(* IEC 61131-3 sources: SortJet_MasterSPS_Aufbau.fbsproj/07_Auftragsverwaltung/BasisSchrittketten, 22 files *)

(* ---- Shuttle_Austransport.fb.st ---- *)
(* METADATA
{
	"v3Meta": {
		"objectGuid": "ac2be6b1-afec-449b-a8c9-7faca61891b0"
	}
}
*)
FUNCTION_BLOCK Shuttle_Austransport
VAR_INPUT

  // BOOLEAN
  bpReset                : BOOL;

  // WORD
  wStation               : WORD;
  wWand                  : WORD;

  // STRUKTUR
  Auftragsdaten          : Auftragsdaten_ST;

END_VAR
VAR_OUTPUT

  // BOOLEAN
  bpDone                 : BOOL;
  bpFehler               : BOOL;

END_VAR
VAR

  // BOOLEAN
  blStationQuittiertScheiben : BOOL;

  // WORD
  wlAustransportstation  : WORD;

  // INT
  ilScheibenZuQuittieren : INT;

  // STEPS
  steplSchritt           : STEPS_TE;

END_VAR
//-------------------------------------------------------------------------------------------------
// STEUERUNG AUSTRANSPORT
//-------------------------------------------------------------------------------------------------
IF ( Auftragsdaten.wAuftrag = eStation_Austransport) THEN

  CASE steplSchritt OF

    // AUSTRANSPORT ===============================================
    STEP_0_E:
      (* Hinweis:
         - Ueberpruefung des Sicherheitskreises
      *)
      IF checkSafetyCircuitsNotBlocked(starrShuttleBasisParameter[wStation]) AND NOT bgShuttleAustransportSperren[wStation]  THEN
        steplSchritt := STEP_10_E;
      END_IF

    // AUSTRANSPORT ===============================================
    STEP_10_E:
      // Auftragsdaten pruefen:
      //  - Sollte es fehler in der Auftragsdatenstruktur geben wird in den Fehlerschritt 900
      //    gesprungen. Die Fehlerauswertung findet in der Funktion Shuttledaten_Pruefen statt.
      steplSchritt := STEP_20_E;

      IF NOT AuftragsdatenPruefen( wStation, wWand, Auftragsdaten) THEN
        steplSchritt := STEP_900_E;
      END_IF

    // AUSTRANSPORT ===============================================
    STEP_20_E:
      // ---------------------------------------------------------------------------------------
      //  AUSTRANSPORT BEDINGUNGEN PRUEFEN
      //
      //  Hinweis:
      // - n/c
      // ---------------------------------------------------------------------------------------

      (* Hinweis:
         - Uebergabe der Quellstation [Sender] fuer den Austransport [Zum ueberpruefen des Zustandes der Station]
      *)
      wlAustransportstation := Auftragsdaten.wTransferstationsNr1;

      starrShuttleBasisParameter[wStation].bRueckwaertsTransportieren[wWand] := FALSE;
      starrShuttleBasisParameter[wStation].bTransferstationTransfershuttle[wWand] := FALSE;

      (* Hinweis:
         - Auftragsdaten ans Shuttle übergeben
      *)
      ilScheibenZuQuittieren :=WORD_TO_INT( Auftragsdaten.wAnzahlScheiben);

      (* Hinweis:
         - Auftragsdaten uebergeben
      *)
      starrShuttleBasisParameter[wStation].pAuftrag[wWand] := Auftragsdaten;

      (* Hinweis:
         - Scheibenführung / Wandverstellung anstellen
         - Aus dem Speicher: Speicherslot dicke nehmen ; von einer Station die Scheibendicke nehmen
      *)
      IF ( starrShuttleBasisParameter[wStation].pAuftrag[wWand].rAuftragsDicke <= wgMKScheibenDicke13mm ) THEN
        starrShuttleBasisParameter[wStation].pAuftrag[wWand].stAuftragsOptionen.eDickenverstellung    := eZylinderStellung16mm;
      ELSIF ( starrShuttleBasisParameter[wStation].pAuftrag[wWand].rAuftragsDicke <= wgMKScheibenDicke19mm ) THEN
        starrShuttleBasisParameter[wStation].pAuftrag[wWand].stAuftragsOptionen.eDickenverstellung    := eZylinderStellung23mm;
      ELSIF ( starrShuttleBasisParameter[wStation].pAuftrag[wWand].rAuftragsDicke <= wgMKScheibenDicke24mm ) THEN
        starrShuttleBasisParameter[wStation].pAuftrag[wWand].stAuftragsOptionen.eDickenverstellung    := eZylinderStellung29mm;
      END_IF

      // Kippen
      starrShuttleBasisParameter[wStation].pAuftrag[wWand].stAuftragsOptionen.eKippen_SollPosition                  := starrShuttleBasisParameter[wStation].stMKs.stSchnittstellendaten.aAustransporte.Kippen[wlAustransportstation];
      starrShuttleBasisParameter[wStation].pAuftrag[wWand].stAuftragsOptionen.eKippen_SollPosition_NachEintransport := 0;
      starrShuttleBasisParameter[wStation].pAuftrag[wWand].stAuftragsOptionen.eKippen_SollPosition_NachAustransport := starrShuttleBasisParameter[wStation].stMKs.stSchnittstellendaten.aAustransporte.KippenNachAustransport[wlAustransportstation];

      // Hub
      starrShuttleBasisParameter[wStation].pAuftrag[wWand].stAuftragsOptionen.eHub                  := starrShuttleBasisParameter[wStation].stMKs.stSchnittstellendaten.aAustransporte.Hub[wlAustransportstation];
      starrShuttleBasisParameter[wStation].pAuftrag[wWand].stAuftragsOptionen.eHub_NachEintransport := 0;
      starrShuttleBasisParameter[wStation].pAuftrag[wWand].stAuftragsOptionen.eHub_NachAustransport := starrShuttleBasisParameter[wStation].stMKs.stSchnittstellendaten.aAustransporte.HubNachAustransport[wlAustransportstation];

      // Greifer [Ausbaustufe stStationsAufbau.bGreifer]: Greiferseite je Partnerstation, Zangenoeffnung wie die Scheibenfuehrung
      starrShuttleBasisParameter[wStation].pAuftrag[wWand].stAuftragsOptionen.eGreiferTyp   := eGreiferDefault;
      IF ( starrShuttleBasisParameter[wStation].stMKs.stStationsAufbau.bGreifer[wWand] ) THEN
        starrShuttleBasisParameter[wStation].pAuftrag[wWand].stAuftragsOptionen.eGreiferTyp := starrShuttleBasisParameter[wStation].stMKs.stSchnittstellendaten.aAustransporte.Greifer[wlAustransportstation];
      END_IF
      starrShuttleBasisParameter[wStation].pAuftrag[wWand].stAuftragsOptionen.eGreiferZangeStellung := starrShuttleBasisParameter[wStation].pAuftrag[wWand].stAuftragsOptionen.eDickenverstellung;

      // Scheibentyp prüfen
      starrShuttleBasisParameter[wStation].wGlasTyp[wWand] := eScheibe_Default;
      IF ( Auftragsdaten.rAuftragsLaenge >= starrShuttleBasisParameter[wStation].stMKs.stStationsParameter.rLaengeUebergroesseScheibe ) THEN
        starrShuttleBasisParameter[wStation].wGlasTyp[wWand] := eScheibe_Maximal;
      END_IF

      (* Hinweis:
         - Stations-Zustand pruefen
      *)
      CASE wlAustransportstation OF

        // Transfershuttles
        cERSTES_TRANSFERSHUTTLE..cLETZTES_TRANSFERSHUTTLE:
          steplSchritt := STEP_200_E;

        // Stationen
        cERSTE_STATION..cLETZTE_STATION:
          IF ( ( Job_Stationen.AuftragsdatenWand[wlAustransportstation, Auftragsdaten.wTransferwand].wAuftrag = eStation_Kein_Auftrag )
               OR ( Job_Stationen.AuftragsdatenWand[wlAustransportstation, Auftragsdaten.wTransferwand].wAuftrag = eStation_Belegt )
               OR ( Job_Stationen.AuftragsdatenWand[wlAustransportstation, Auftragsdaten.wTransferwand].wAuftrag = eStation_Durchtransport ) )
          THEN
            steplSchritt := STEP_100_E;
          END_IF

        cERSTE_FREMDANLAGE_AUSLAUF..cLETZTE_FREMDANLAGE_AUSLAUF:
          IF ( Auftragsdaten.wTransferstationsNr2 <> 0 ) THEN
            IF   ( Job_Fremdanlage.AuftragsdatenFremdanlage[wlAustransportstation].wAuftrag = eStation_Kein_Auftrag )
                 AND ( Job_Stationen.AuftragsdatenWand[Auftragsdaten.wTransferstationsNr2, Auftragsdaten.wTransferwand].wAuftrag = eStation_Kein_Auftrag )
            THEN
              steplSchritt := STEP_100_E;
            END_IF
          ELSE
            IF ( Job_Fremdanlage.AuftragsdatenFremdanlage[wlAustransportstation].wAuftrag = eStation_Kein_Auftrag )
            THEN
              steplSchritt := STEP_100_E;
            END_IF
          END_IF

        // Fremdanlage
        cERSTE_FREMDANLAGE_EINLAUF..cLETZTE_FREMDANLAGE_EINLAUF:
          ;

        // Faecherwagen direkt (Transferstation 1): nur mit dem Greifer. Ohne Greifer geht es in den Faecherwagen ueber ein
        // Transfershuttle mit bTransferShuttleFuerFaecherwagen (Transferstation 1 = Transfershuttle, Transferstation 2 = Faecherwagen)
        cERSTE_FAECHERWAGENSTATIONS_NR..cLETZTE_FAECHERWAGENSTATIONS_NR:
          IF ( starrShuttleBasisParameter[wStation].pAuftrag[wWand].stAuftragsOptionen.eGreiferTyp <> eGreiferDefault ) THEN
            IF ( starrFaecherwagenBasisParameter[wlAustransportstation].OutGlasTransport[cWAND_1].bBereitZumEintransport ) THEN
              steplSchritt := STEP_100_E;
            END_IF
          ELSE
            wpgFehlerdaten[0] := starrShuttleBasisParameter[wStation].stMKs.stStationsNummern.NummerExtern;
            wpgFehlerdaten[1] := wWand;
            SpsError( eFehler_Station,
                      cMELDUNG_AUFTRAGSDATEN_FALSCHE_AUSLAUFSTATION,
                      starrShuttleBasisParameter[wStation].stMKs.stStationsNummern.NummerIntern,
                      AutomatikkreisBestimmen(starrShuttleBasisParameter[wStation].stMKs.stStationsNummern.NummerSPS),
                      wpgFehlerdaten );

            steplSchritt := STEP_900_E;
          END_IF

        ELSE
          wpgFehlerdaten[0] := starrShuttleBasisParameter[wStation].stMKs.stStationsNummern.NummerExtern;
          wpgFehlerdaten[1] := wWand;
          SpsError( eFehler_Station,
                    cMELDUNG_AUFTRAGSDATEN_FALSCHE_AUSLAUFSTATION,
                    starrShuttleBasisParameter[wStation].stMKs.stStationsNummern.NummerIntern,
                    AutomatikkreisBestimmen(starrShuttleBasisParameter[wStation].stMKs.stStationsNummern.NummerSPS),
                    wpgFehlerdaten );

          steplSchritt := STEP_900_E;

      END_CASE

    // AUSTRANSPORT ==============================================
    STEP_100_E:
      (* Hinweis:
         - Auftrag ab Station übergeben und Shuttle Informationen zuweisen
      *)
      CASE wlAustransportstation OF

        // Stationen
        cERSTE_STATION..cLETZTE_STATION:

          IF AutomatikAktiv(wlAustransportstation) THEN

            (* Hinweis:
               - Auftragsdaten in Transferstation kopieren
            *)
            IF NOT ( Job_Stationen.AuftragsdatenWand[wlAustransportstation, Auftragsdaten.wTransferwand].wAuftrag = eStation_Durchtransport ) THEN
              Job_Stationen.AuftragsdatenWand[wlAustransportstation, Auftragsdaten.wTransferwand]           := AuftragsdatenUmkopieren(FALSE, FALSE, Auftragsdaten);
              Job_Stationen.AuftragsdatenWand[wlAustransportstation, Auftragsdaten.wTransferwand].wAuftrag  := eStation_Eintransport;
            END_IF

            (* Hinweis:
               - Kopplung zur Transferstation herstellen
            *)
            starrShuttleBasisParameter[wStation].InGlasTransportNachfolger[wWand] := starrStationBasisParameter[wlAustransportstation].OutGlasTransport[Auftragsdaten.wTransferwand];
            starrShuttleBasisParameter[wStation].InGlasTransportVorgaenger[wWand] := starrStationBasisParameter[wlAustransportstation].OutGlasTransport[Auftragsdaten.wTransferwand];

            (* Hinweis:
               - Daten an das Shuttle uebergeben
            *)
            starrShuttleBasisParameter[wStation].bAustransport[wWand]                  := TRUE;
            starrShuttleBasisParameter[wStation].bRueckwaertsTransportieren[wWand]     := ( starrShuttleBasisParameter[wStation].stMKs.stSchnittstellendaten.aAustransporte.Station[wlAustransportstation] = Rueckwaertig );

            steplSchritt := STEP_400_E;

          END_IF

        cERSTE_FREMDANLAGE_AUSLAUF..cLETZTE_FREMDANLAGE_AUSLAUF:

          IF ( Auftragsdaten.wTransferstationsNr2 <> 0 ) THEN

            IF AutomatikAktiv(Auftragsdaten.wTransferstationsNr2) THEN

              (* Hinweis:
                 - Kopplung zur Transferstation herstellen
              *)
              starrShuttleBasisParameter[wStation].InGlasTransportNachfolger[wWand] := starrStationBasisParameter[Auftragsdaten.wTransferstationsNr2].OutGlasTransport[Auftragsdaten.wTransferwand];
              starrShuttleBasisParameter[wStation].InGlasTransportVorgaenger[wWand] := starrStationBasisParameter[Auftragsdaten.wTransferstationsNr2].OutGlasTransport[Auftragsdaten.wTransferwand];

              (* Hinweis:
                 - Auftragsdaten in Transferstation kopieren
              *)
              Job_Fremdanlage.AuftragsdatenFremdanlage[wlAustransportstation]          := AuftragsdatenUmkopieren(FALSE, FALSE, Auftragsdaten);
              Job_Fremdanlage.AuftragsdatenFremdanlage[wlAustransportstation].wAuftrag := eStation_Eintransport;

              (* Hinweis:
                 - Daten an das Shuttle uebergeben
              *)
              starrShuttleBasisParameter[wStation].bAustransport[wWand]                  := TRUE;
              starrShuttleBasisParameter[wStation].bRueckwaertsTransportieren[wWand]     := ( starrShuttleBasisParameter[wStation].stMKs.stSchnittstellendaten.aAustransporte.Station[wlAustransportstation] = Rueckwaertig );

              steplSchritt := STEP_400_E;

            END_IF

          ELSE

            (* Hinweis:
               - Kopplung zur Transferstation herstellen
            *)
            starrShuttleBasisParameter[wStation].InGlasTransportNachfolger[wWand] := starrFremdanlageAuslaufStationBasisParameter[wlAustransportstation].OutGlasTransport[cWAND_1];
            starrShuttleBasisParameter[wStation].InGlasTransportVorgaenger[wWand] := starrFremdanlageAuslaufStationBasisParameter[wlAustransportstation].OutGlasTransport[cWAND_1];
            starrFremdanlageAuslaufStationBasisParameter[wlAustransportstation].InGlasTransportVorgaenger[cWAND_1] :=  starrShuttleBasisParameter[wStation].OutGlasTransport[wWand];

            (* Hinweis:
               - Auftragsdaten in Transferstation kopieren
            *)
            Job_Fremdanlage.AuftragsdatenFremdanlage[wlAustransportstation]          := AuftragsdatenUmkopieren(FALSE, FALSE, Auftragsdaten);
            Job_Fremdanlage.AuftragsdatenFremdanlage[wlAustransportstation].wAuftrag := eStation_Eintransport;

            (* Hinweis:
               - Daten an das Shuttle uebergeben
            *)
            starrShuttleBasisParameter[wStation].bAustransport[wWand]              := TRUE;
            starrShuttleBasisParameter[wStation].bRueckwaertsTransportieren[wWand] := ( starrShuttleBasisParameter[wStation].stMKs.stSchnittstellendaten.aAustransporte.Station[wlAustransportstation] = Rueckwaertig );

            steplSchritt := STEP_400_E;

          END_IF

        cERSTE_FAECHERWAGENSTATIONS_NR..cLETZTE_FAECHERWAGENSTATIONS_NR:
          (* Hinweis:
             - Austransport in den Faecherwagen mit dem Greifer (Greiferseite im Auftrag)
          *)
          starrShuttleBasisParameter[wStation].bRueckwaertsTransportieren[wWand] := FALSE;
          starrShuttleBasisParameter[wStation].bAustransport[wWand]              := TRUE;

          steplSchritt := STEP_400_E;

      END_CASE

    // AUSTRANSPORT ===============================================
    STEP_200_E:
      // ---------------------------------------------------------------------------------------
      //  EINTRANSPORT MITTELS TRANSFERSHUTTLE
      //
      //  Hinweis:
      //  - Transferstation2 = 0   => Eintransport mit nur einem Transfershuttle
      //  - Transferstation2 <> 0  => Eintransport im Transfershuttle-Verbund
      // ---------------------------------------------------------------------------------------

      IF ( Auftragsdaten.wTransferstationsNr2 = 0 OR starrTransfershuttleBasisParameter[wlAustransportstation].stMKs.stStationsOptionen.stTransfershuttle.bTransferShuttleFuerFaecherwagen ) THEN

        IF (  ( Job_Shuttle.AuftragsdatenTransfershuttle[wlAustransportstation].wAuftrag = eStation_Kein_Auftrag ) ) THEN
          steplSchritt := STEP_210_E;
        END_IF

      ELSE
        VailiderenTransfershuttleVerbund ( wTransferstation1 := wlAustransportstation,
                                           wTransferstation2 := Auftragsdaten.wTransferstationsNr2 );

        IF (  ( Job_Shuttle.AuftragsdatenTransfershuttle[wlAustransportstation].wAuftrag = eStation_Kein_Auftrag )
             AND ( Job_Shuttle.AuftragsdatenTransfershuttle[Auftragsdaten.wTransferstationsNr2].wAuftrag  = eStation_Kein_Auftrag ) )
        THEN
          steplSchritt := STEP_220_E;
        END_IF

      END_IF

    // AUSTRANSPORT ===============================================
    STEP_210_E:
      // ---------------------------------------------------------------------------------------
      //  EINTRANSPORT TRANSFERSHUTTLE [DEFAULT]
      //
      //  Hinweis:
      // - n/c
      // ---------------------------------------------------------------------------------------

      (* Hinweis:
         - Kopplung
      *)
      IF ( starrShuttleBasisParameter[wStation].stMKs.stSchnittstellendaten.aAustransporte.Station[wlAustransportstation] = Rueckwaertig ) THEN
        starrTransfershuttleBasisParameter[wlAustransportstation].InGlasTransportNachfolger[wWand] := starrShuttleBasisParameter[wStation].OutGlasTransport[wWand];
        starrShuttleBasisParameter[wStation].InGlasTransportVorgaenger[wWand] := starrTransfershuttleBasisParameter[wlAustransportstation].OutGlasTransport[wWand];

      ELSE
        starrTransfershuttleBasisParameter[wlAustransportstation].InGlasTransportVorgaenger[wWand] := starrShuttleBasisParameter[wStation].OutGlasTransport[wWand];
        starrShuttleBasisParameter[wStation].InGlasTransportNachfolger[wWand] := starrTransfershuttleBasisParameter[wlAustransportstation].OutGlasTransport[wWand];

      END_IF

      (* Hinweis:
         - TS auf FW koppeln
      *)
      IF   starrTransfershuttleBasisParameter[wlAustransportstation].stMKs.stStationsOptionen.stTransfershuttle.bTransferShuttleFuerFaecherwagen
           AND IsBetweenWORD(Auftragsdaten.wTransferstationsNr2, cERSTE_FAECHERWAGENSTATIONS_NR, cLETZTE_FAECHERWAGENSTATIONS_NR)
      THEN
        IF ( starrShuttleBasisParameter[wStation].stMKs.stSchnittstellendaten.aAustransporte.Station[wlAustransportstation] = Rueckwaertig ) THEN
          starrTransfershuttleBasisParameter[wlAustransportstation].InGlasTransportVorgaenger[wWand] := starrFaecherwagenBasisParameter[Auftragsdaten.wTransferstationsNr2].OutGlasTransport[cWAND_1];
        ELSE
          starrTransfershuttleBasisParameter[wlAustransportstation].InGlasTransportNachfolger[wWand] := starrFaecherwagenBasisParameter[Auftragsdaten.wTransferstationsNr2].OutGlasTransport[cWAND_1];
        END_IF
      END_IF

      (* Hinweis:
         - Neuen Auftag in den FIFO [Warteschlange] eintragen
      *)
      Job_Shuttle.AuftragsdatenTransfershuttle[wlAustransportstation]          := AuftragsdatenUmkopieren(FALSE, FALSE, Auftragsdaten);
      Job_Shuttle.AuftragsdatenTransfershuttle[wlAustransportstation].wAuftrag := eStation_Eintransport;

      starrShuttleBasisParameter[wStation].bScheibentrennen[wWand]                := FALSE;
      starrShuttleBasisParameter[wStation].bRueckwaertsTransportieren[wWand]      := ( starrShuttleBasisParameter[wStation].stMKs.stSchnittstellendaten.aAustransporte.Station[wlAustransportstation] = Rueckwaertig );
      starrShuttleBasisParameter[wStation].bAustransport[wWand]                   := TRUE;
      starrShuttleBasisParameter[wStation].bTransferstationTransfershuttle[wWand] := TRUE;

      steplSchritt := STEP_400_E;

    // AUSTRANSPORT ===============================================
    STEP_220_E:
      // ---------------------------------------------------------------------------------------
      //  EINTRANSPORT TRANSFERSHUTTLE [VERBUND]
      //
      //  Hinweis:
      //  - n/c
      // ---------------------------------------------------------------------------------------

      (* Hinweis:
         - Kopplung
      *)
      IF ( starrShuttleBasisParameter[wStation].stMKs.eStationsTyp = eInputshuttle ) THEN
        starrTransfershuttleBasisParameter[wlAustransportstation].InGlasTransportVorgaenger[wWand] := starrShuttleBasisParameter[wStation].OutGlasTransport[wWand];
        starrShuttleBasisParameter[wStation].InGlasTransportNachfolger[wWand] := starrTransfershuttleBasisParameter[wlAustransportstation].OutGlasTransport[wWand];

      ELSE
        starrTransfershuttleBasisParameter[wlAustransportstation].InGlasTransportNachfolger[wWand] := starrShuttleBasisParameter[wStation].OutGlasTransport[wWand];
        starrShuttleBasisParameter[wStation].InGlasTransportVorgaenger[wWand] := starrTransfershuttleBasisParameter[wlAustransportstation].OutGlasTransport[wWand];

      END_IF

      (* Hinweis:
         - Transfershuttle koppeln
      *)
      aTransfershuttles[wlAustransportstation].stpInTransportVerbund  := aTransfershuttles[Auftragsdaten.wTransferstationsNr2].stpOutTransportVerbund;
      aTransfershuttles[Auftragsdaten.wTransferstationsNr2].stpInTransportVerbund   := aTransfershuttles[wlAustransportstation].stpOutTransportVerbund;

      (* Hinweis:
         - Auftragsdaten an die Transfershuttle uebergeben
      *)
      Job_Shuttle.AuftragsdatenTransfershuttle[wlAustransportstation]          := AuftragsdatenUmkopieren(FALSE, FALSE, Auftragsdaten);
      Job_Shuttle.AuftragsdatenTransfershuttle[wlAustransportstation].wAuftrag := eStation_Eintransport;

      Job_Shuttle.AuftragsdatenTransfershuttle[Auftragsdaten.wTransferstationsNr2]           := AuftragsdatenUmkopieren(TRUE, FALSE, Auftragsdaten);
      Job_Shuttle.AuftragsdatenTransfershuttle[Auftragsdaten.wTransferstationsNr2].wAuftrag  := eStation_Transportkopplung;

      starrShuttleBasisParameter[wStation].bScheibentrennen[wWand]                := FALSE;
      starrShuttleBasisParameter[wStation].bRueckwaertsTransportieren[wWand]      := ( starrShuttleBasisParameter[wStation].stMKs.stSchnittstellendaten.aAustransporte.Station[wlAustransportstation] = Rueckwaertig );
      starrShuttleBasisParameter[wStation].bAustransport[wWand]                   := TRUE;
      starrShuttleBasisParameter[wStation].bTransferstationTransfershuttle[wWand] := TRUE;

      steplSchritt := STEP_400_E;

    // AUSTRANSPORT ===============================================
    STEP_400_E:
      // ---------------------------------------------------------------------------------------
      //  QUITTIERUNGEN UND EINTRANSPORT- ABSCHLUSS
      //
      //  Hinweis:
      //  - Scheibenquittieren: Message zur MMI
      // ---------------------------------------------------------------------------------------
      blStationQuittiertScheiben := starrShuttleBasisParameter[wStation].stMKs.stSchnittstellendaten.aAustransporte.bStationQuittiertScheibe[wlAustransportstation];

      IF ( starrShuttleBasisParameter[wStation].OutGlasTransport[wWand].bQuittScheibe ) THEN

        IF ( ilScheibenZuQuittieren > 0 ) THEN

          wSps2MmiZielStation  := Auftragsdaten.wTransferstationsNr1;
          wSps2MmiQuellStation := starrShuttleBasisParameter[wStation].stMKs.stStationsNummern.NummerIntern;
          wSps2MmiZielWand     := Auftragsdaten.wTransferwand;
          wSps2MmiQuellWand    := wWand;
          dwSps2MmiWartezeit   := starrShuttleBasisParameter[wStation].dwWartezeit[wWand];
          wSPS2MMIAuftragstyp  := 1;

          MsgToMmi(auftragsnr_w := SB0_SPS_QUIT_SHEET_ORDER );
        END_IF

        ilScheibenZuQuittieren := ilScheibenZuQuittieren - 1;

      END_IF

      (* Hinweis:
         - Abschliessen des Austransports
      *)
      IF ( starrShuttleBasisParameter[wStation].bAustransportAbgeschlossen[wWand] ) THEN

        starrShuttleBasisParameter[wStation].bAustransport[wWand]                 := FALSE;
        starrShuttleBasisParameter[wStation].bRueckwaertsTransportieren[wWand]    := FALSE;

        steplSchritt := STEP_410_E;
      END_IF

      (* Fehlerbehandlung:
         - Inputshuttle
      *)
      IF ( starrShuttleBasisParameter[wStation].bFehler ) THEN
        SpsError( eFehler_Station,
                  starrShuttleBasisParameter[wStation].wFehlerNummer,
                  starrShuttleBasisParameter[wStation].stMKs.stStationsNummern.NummerIntern,
                  AutomatikkreisBestimmen(starrShuttleBasisParameter[wStation].stMKs.stStationsNummern.NummerSPS),
                  starrShuttleBasisParameter[wStation].awFehlerInformationen );

        steplSchritt := STEP_900_E;
      END_IF

    // AUSTRANSPORT ==============================================
    STEP_410_E:
      (* Anmerkung:
         - Gueltige Anzahl von Scheiben wurden quittiert
      *)
      IF ( ilScheibenZuQuittieren = 0 ) THEN
        steplSchritt := STEP_1000_E;

      (* Anmerkung:
         - Zu wenig Scheiben quittiert
      *)
      ELSIF ( ilScheibenZuQuittieren > 0 ) THEN
        wpgFehlerdaten[0] := starrShuttleBasisParameter[wStation].stMKs.stStationsNummern.NummerExtern;
        wpgFehlerdaten[1] := wWand;

        SpsError( eFehler_Station,
                  cMELDUNG_STATION_ZUWENIG_SCHEIBEN_QUITTIERT_WAND_AUSTRANSPORT,
                  starrShuttleBasisParameter[wStation].stMKs.stStationsNummern.NummerIntern,
                  AutomatikkreisBestimmen(starrShuttleBasisParameter[wStation].stMKs.stStationsNummern.NummerSPS),
                  wpgFehlerdaten );

        steplSchritt := STEP_900_E;

      (* Anmerkung:
         - Zu viele Scheiben quittiert
      *)
      ELSIF ( ilScheibenZuQuittieren < 0 ) THEN
        wpgFehlerdaten[0] := starrShuttleBasisParameter[wStation].stMKs.stStationsNummern.NummerExtern;
        wpgFehlerdaten[1] := wWand;

        SpsError( eFehler_Station,
                  cMELDUNG_STATION_ZUVIELE_SCHEIBEN_QUITTIERT_WAND_AUSTRANSPORT,
                  starrShuttleBasisParameter[wStation].stMKs.stStationsNummern.NummerIntern,
                  AutomatikkreisBestimmen(starrShuttleBasisParameter[wStation].stMKs.stStationsNummern.NummerSPS),
                  wpgFehlerdaten );

        steplSchritt := STEP_900_E;
      END_IF

    // AUSTRANSPORT ===============================================
    STEP_900_E:
      bpFehler := TRUE;

    // AUSTRANSPORT ===============================================
    STEP_1000_E:
      bpDone := TRUE;
      Auftragsdaten.wAuftrag := eStation_Kein_Auftrag;

  // AUSTRANSPORT ===============================================
  END_CASE

END_IF

IF bpReset THEN
  bpFehler := FALSE;
  bpDone := FALSE;
  bpReset := FALSE;
  starrShuttleBasisParameter[wStation].bAustransport[wWand] := FALSE;
  starrShuttleBasisParameter[wStation].bTransferstationTransfershuttle[wWand] := FALSE;
  steplSchritt := STEP_0_E;
END_IF
END_FUNCTION_BLOCK

(* ---- Shuttle_Durchtransport.fb.st ---- *)
(* METADATA
{
	"v3Meta": {
		"objectGuid": "d20ae107-ce5b-4166-b2bd-9e4de3a442ef"
	}
}
*)
FUNCTION_BLOCK Shuttle_Durchtransport
VAR_INPUT

  // BOOLEAN
  bpReset                : BOOL;

  // WORD
  wStation               : WORD;
  wWand                  : WORD;

  // STRUKTUR
  Auftragsdaten          : Auftragsdaten_ST;

END_VAR
VAR_OUTPUT

  // BOOLEAN
  bpDone                 : BOOL;
  bpFehler               : BOOL;

END_VAR
VAR

  // BOOLEAN
  blStationQuittiertScheiben             : BOOL;
  blKopplungGefundenEintransport         : BOOL;
  blKopplungGefundenAustransport         : BOOL;

  // WORD
  wlEintransportstation : WORD;
  wlAustransportstation : WORD;

  // INT
  ilScheibenZuQuittieren : INT;

  // STEPS
  steplSchritt           : STEPS_TE;

END_VAR

//-------------------------------------------------------------------------------------------------
// STEUERUNG DURCHTRANSPORT
//-------------------------------------------------------------------------------------------------
IF Auftragsdaten.wAuftrag = eStation_Durchtransport THEN
  CASE steplSchritt OF
    // DURCHTRANSPORT =================================
    STEP_0_E:
      (* Hinweis:
         - Ueberpruefung des Sicherheitskreises
      *)
      IF checkSafetyCircuitsNotBlocked(starrShuttleBasisParameter[wStation]) AND NOT bgShuttleEintransportSperren[wStation] AND NOT bgShuttleAustransportSperren[wStation]  THEN
        steplSchritt := STEP_10_E;
      END_IF

    // DURCHTRANSPORT ==================================================
    STEP_10_E:
      // Auftragsdaten pruefen:
      //  - Sollte es fehler in der Auftragsdatenstruktur geben wird in den Fehlerschritt 900
      //    gesprungen. Die Fehlerauswertung findet in der Funktion Shuttledaten_Pruefen statt.
      steplSchritt := STEP_20_E;

      IF NOT AuftragsdatenPruefen( wStation, wWand, Auftragsdaten) THEN
        steplSchritt := STEP_900_E;
      END_IF

    // DURCHTRANSPORT =================================
    STEP_20_E:
      (* Hinweis:
         - Kopplung fuer diesen Auftrag neu bestimmen. Sonst ueberschreibt ein Merker aus dem letzten Auftrag den Fehlerschritt.
      *)
      blKopplungGefundenEintransport := FALSE;
      blKopplungGefundenAustransport := FALSE;

      (* Hinweis:
         - Uebergabe der Quellstation [Sender] fuer den Austransport [Zum ueberpruefen des Zustandes der Station]
      *)
      wlEintransportstation := Auftragsdaten.wTransferstationsNr1;
      wlAustransportstation := Auftragsdaten.wTransferstationsNr2;

      (* Hinweis:
         - Zuweisung Transportkopplung
      *)
      CASE wlEintransportstation OF

        // Stationen
        cERSTE_STATION..cLETZTE_STATION:
          (* Hinweis:
             - Transportkopplung
          *)
          IF ( starrShuttleBasisParameter[wStation].stMKs.stSchnittstellendaten.aEintransporte.Station[wlEintransportstation] = Vorwaertig ) THEN
            starrShuttleBasisParameter[wStation].InGlasTransportVorgaenger[wWand] := starrStationBasisParameter[wlEintransportstation].OutGlasTransport[Auftragsdaten.wTransferwand];
          ELSE
            starrShuttleBasisParameter[wStation].InGlasTransportNachfolger[wWand] := starrStationBasisParameter[wlEintransportstation].OutGlasTransport[Auftragsdaten.wTransferwand];
          END_IF
          blKopplungGefundenEintransport := TRUE;

        ELSE
          wpgFehlerdaten[0] := starrShuttleBasisParameter[wStation].stMKs.stStationsNummern.NummerExtern;
          wpgFehlerdaten[1] := wlEintransportstation;
          SpsError( eFehler_Station,
                    cMELDUNG_AUFTRAGSDATEN_FALSCHE_EINLAUFSTATION,
                    starrShuttleBasisParameter[wStation].stMKs.stStationsNummern.NummerIntern,
                    AutomatikkreisBestimmen(starrShuttleBasisParameter[wStation].stMKs.stStationsNummern.NummerSPS),
                    wpgFehlerdaten );

          steplSchritt := STEP_900_E;

      END_CASE

      (* Hinweis:
         - Zuweisung Transportkopplung
      *)
      CASE wlAustransportstation OF

        // Stationen
        cERSTE_STATION..cLETZTE_STATION:
          (* Hinweis:
             - Transportkopplung
          *)
          IF ( starrShuttleBasisParameter[wStation].stMKs.stSchnittstellendaten.aAustransporte.Station[wlAustransportstation] = Vorwaertig ) THEN
            starrShuttleBasisParameter[wStation].InGlasTransportNachfolger[wWand] := starrStationBasisParameter[wlAustransportstation].OutGlasTransport[Auftragsdaten.wTransferwand];
          ELSE
            starrShuttleBasisParameter[wStation].InGlasTransportVorgaenger[wWand] := starrStationBasisParameter[wlAustransportstation].OutGlasTransport[Auftragsdaten.wTransferwand];
          END_IF
          blKopplungGefundenAustransport := TRUE;

        cERSTE_FREMDANLAGE_AUSLAUF..cLETZTE_FREMDANLAGE_AUSLAUF:
          (* Hinweis:
             - Transportkopplung
          *)
          IF ( starrShuttleBasisParameter[wStation].stMKs.stSchnittstellendaten.aAustransporte.Station[wlAustransportstation] = Vorwaertig ) THEN
            starrShuttleBasisParameter[wStation].InGlasTransportNachfolger[wWand] := starrFremdanlageAuslaufStationBasisParameter[wlAustransportstation].OutGlasTransport[cWAND_1];
          ELSE
            starrShuttleBasisParameter[wStation].InGlasTransportVorgaenger[wWand] := starrFremdanlageAuslaufStationBasisParameter[wlAustransportstation].OutGlasTransport[cWAND_1];
          END_IF
          blKopplungGefundenAustransport := TRUE;

        ELSE
          wpgFehlerdaten[0] := starrShuttleBasisParameter[wStation].stMKs.stStationsNummern.NummerExtern;
          wpgFehlerdaten[1] := wlAustransportstation;
          SpsError( eFehler_Station,
                    cMELDUNG_AUFTRAGSDATEN_FALSCHE_AUSLAUFSTATION,
                    starrShuttleBasisParameter[wStation].stMKs.stStationsNummern.NummerIntern,
                    AutomatikkreisBestimmen(starrShuttleBasisParameter[wStation].stMKs.stStationsNummern.NummerSPS),
                    wpgFehlerdaten );

          steplSchritt := STEP_900_E;

      END_CASE

      IF blKopplungGefundenEintransport AND blKopplungGefundenAustransport THEN
        steplSchritt := STEP_30_E;
      END_IF

    // DURCHTRANSPORT =================================
    STEP_30_E:

      (* Hinweis:
         - Scheibenquittierung
      *)
      ilScheibenZuQuittieren := WORD_TO_INT(Auftragsdaten.wAnzahlScheiben);

      (* Hinweis:
         - Auftrags- Optionen bestimmen und zuweisen
      *)
      Auftragsdaten.stAuftragsOptionen.eKippen_SollPosition := starrShuttleBasisParameter[wStation].stMKs.stSchnittstellendaten.aEintransporte.Kippen[wlEintransportstation];

      IF ( Auftragsdaten.rAuftragsDicke < wgUnterteilerMinMaxGlasdicke ) THEN
        Auftragsdaten.stAuftragsOptionen.eDickenverstellung := eZylinderStellung16mm;
      ELSE
        Auftragsdaten.stAuftragsOptionen.eDickenverstellung := eZylinderStellung23mm;
      END_IF
      Auftragsdaten.stAuftragsOptionen.eDrehen_Sollposition := 0;
      Auftragsdaten.stAuftragsOptionen.eDrehen_Sollposition_NachAustransport := 0;
      Auftragsdaten.stAuftragsOptionen.eKippen_SollPosition_NachAustransport := 0;
      Auftragsdaten.stAuftragsOptionen.eGlastransport := 0;
      Auftragsdaten.stAuftragsOptionen.eHub                  := starrShuttleBasisParameter[wStation].stMKs.stSchnittstellendaten.aEintransporte.Hub[wlEintransportstation];
      Auftragsdaten.stAuftragsOptionen.eHub_NachEintransport := 0;
      Auftragsdaten.stAuftragsOptionen.eHub_NachAustransport := 0;
      Auftragsdaten.stAuftragsOptionen.eQuerachse := 0;
      Auftragsdaten.stAuftragsOptionen.eAchsrichtung := 0;
      Auftragsdaten.stAuftragsOptionen.wMaxTransportGeschwindigkeit:= 0;
      Auftragsdaten.stAuftragsOptionen.eDrehen_Sollposition_NachEintransport := 0;
      Auftragsdaten.stAuftragsOptionen.eKippen_SollPosition_NachEintransport := 0;

      (* Hinweis:
         - Auftragsdaten zuweisen und Eintransport der Station starten
      *)
      starrShuttleBasisParameter[wStation].pAuftrag[wWand] := Auftragsdaten;

      starrShuttleBasisParameter[wStation].bScheibentrennen[wWand]           := FALSE;
      starrShuttleBasisParameter[wStation].bRueckwaertsTransportieren[wWand] := ( starrShuttleBasisParameter[wStation].stMKs.stSchnittstellendaten.aEintransporte.Station[wlEintransportstation] = Rueckwaertig )
                                                                                AND ( starrShuttleBasisParameter[wStation].stMKs.stSchnittstellendaten.aAustransporte.Station[wlAustransportstation] = Rueckwaertig );
      starrShuttleBasisParameter[wStation].bDurchtransport[wWand]            := TRUE;

      steplSchritt := STEP_40_E;

    // AUSTRANSPORT =================================
    STEP_40_E:

      (* Hinweis:
         - Scheibenzaehler dekrementieren
         - Scheibe quittieren, sofern dies nötig ist
      *)
      blStationQuittiertScheiben := starrShuttleBasisParameter[wStation].stMKs.stSchnittstellendaten.aEintransporte.bStationQuittiertScheibe[wlEintransportstation];

      IF ( starrShuttleBasisParameter[wStation].OutGlasTransport[wWand].bQuittScheibe ) THEN

        IF ( ilScheibenZuQuittieren > 0 ) AND blStationQuittiertScheiben THEN

          wSps2MmiZielStation  := starrShuttleBasisParameter[wStation].stMKs.stStationsNummern.NummerIntern;
          wSps2MmiQuellStation := wlEintransportstation;
          wSps2MmiZielWand     := Auftragsdaten.wStationsWand;
          wSps2MmiQuellWand    := Auftragsdaten.wTransferwand;
          dwSps2MmiWartezeit   := starrShuttleBasisParameter[wStation].dwWartezeit[wWand];
          wSPS2MMIAuftragstyp  := 0;

          MsgToMmi(auftragsnr_w := SB0_SPS_QUIT_SHEET_ORDER );

        END_IF

        ilScheibenZuQuittieren := ilScheibenZuQuittieren - 1;

      END_IF

      (* Hinweis:
         - Abschliessen des Austransport
      *)
      IF ( starrShuttleBasisParameter[wStation].bDurchtransportAbgeschlossen[wWand] ) THEN
        starrShuttleBasisParameter[wStation].bRueckwaertsTransportieren[wWand] := FALSE;
        starrShuttleBasisParameter[wStation].bDurchtransport[wWand] := FALSE;
        steplSchritt := STEP_1000_E;
      END_IF

      (* Fehlerbehandlung:
         - Station
      *)
      IF ( starrShuttleBasisParameter[wStation].bFehler ) THEN
        SpsError( eFehler_Station,
                  starrShuttleBasisParameter[wStation].wFehlerNummer,
                  starrShuttleBasisParameter[wStation].stMKs.stStationsNummern.NummerIntern,
                  AutomatikkreisBestimmen(starrShuttleBasisParameter[wStation].stMKs.stStationsNummern.NummerSPS),
                  starrShuttleBasisParameter[wStation].awFehlerInformationen );

        starrShuttleBasisParameter[wStation].bDurchtransport[wWand] := FALSE;
        starrShuttleBasisParameter[wStation].bRueckwaertsTransportieren[wWand] := FALSE;
        steplSchritt := STEP_900_E;
      END_IF

    // DURCHTRANSPORT =================================
    STEP_900_E:
      bpFehler := TRUE;

    // DURCHTRANSPORT =================================
    STEP_1000_E:
      bpDone := TRUE;
      Auftragsdaten.wAuftrag := eStation_Kein_Auftrag;

  END_CASE

END_IF

IF bpReset THEN
  bpFehler := FALSE;
  bpReset := FALSE;
  bpDone := FALSE;
  blKopplungGefundenEintransport := FALSE;
  blKopplungGefundenAustransport := FALSE;
  steplSchritt := STEP_0_E;
  starrShuttleBasisParameter[wStation].bRueckwaertsTransportieren[wWand] := FALSE;
  starrShuttleBasisParameter[wStation].bDurchtransport[wWand] := FALSE;
END_IF
END_FUNCTION_BLOCK

(* ---- Shuttle_Eintransport.fb.st ---- *)
(* METADATA
{
	"v3Meta": {
		"objectGuid": "07a4896b-4b10-421b-8c15-d73c62ab9e42"
	}
}
*)
FUNCTION_BLOCK Shuttle_Eintransport
VAR_INPUT

  // BOOLEAN
  bpReset                : BOOL;

  // WORD
  wStation               : WORD;
  wWand                  : WORD;

  // STRUKTUR
  Auftragsdaten          : Auftragsdaten_ST;

END_VAR
VAR_OUTPUT

  // BOOLEAN
  bpDone                 : BOOL;
  bpFehler               : BOOL;

END_VAR
VAR

  // BOOLEAN
  blStationQuittiertScheiben : BOOL;

  // WORD
  wlEintransportstation  : WORD;

  // INT
  ilScheibenZuQuittieren : INT;

  // STEPS
  steplSchritt           : STEPS_TE;

END_VAR

//-------------------------------------------------------------------------------------------------
// STEUERUNG EINTRANSPORT
//-------------------------------------------------------------------------------------------------
IF ( Auftragsdaten.wAuftrag = eStation_Eintransport ) THEN

  CASE steplSchritt OF

    // EINTRANSPORT ==============================================
    STEP_0_E:
      (* Hinweis:
         - Ueberpruefung des Sicherheitskreises
      *)
      IF checkSafetyCircuitsNotBlocked(starrShuttleBasisParameter[wStation]) AND NOT bgShuttleEintransportSperren[wStation] THEN
        steplSchritt := STEP_10_E;
      END_IF

    // EINTRANSPORT ==============================================
    STEP_10_E:
      // Auftragsdaten pruefen:
      //   - Sollte es fehler in der Auftragsdatenstruktur geben wird in den Fehlerschritt 900
      //   - gesprungen. Die Fehlerauswertung findet in der Funktion Shuttledaten_Pruefen statt.
      steplSchritt := STEP_20_E;

      IF NOT AuftragsdatenPruefen( wStation, wWand, Auftragsdaten) THEN
        steplSchritt := STEP_900_E;
      END_IF

    // EINTRANSPORT ==============================================
    STEP_20_E:
      (* Hinweis:
         - Uebergabe der Quellstation [Sender] fuer den Austransport [Zum ueberpruefen des Zustandes der Station]
      *)
      wlEintransportstation := Auftragsdaten.wTransferstationsNr1;

      starrShuttleBasisParameter[wStation].bRueckwaertsTransportieren[wWand] := FALSE;
      starrShuttleBasisParameter[wStation].bTransferstationTransfershuttle[wWand] := FALSE;

      (* Hinweis:
         - Auftragsdaten ans Shuttle übergeben
      *)
      ilScheibenZuQuittieren := WORD_TO_INT( Auftragsdaten.wAnzahlScheiben );

      (* Hinweis:
         - Auftragsdaten uebergeben
      *)
      starrShuttleBasisParameter[wStation].pAuftrag[wWand] := Auftragsdaten;

      (* Hinweis:
         - Scheibenführung / Wandverstellung anstellen
         - Aus dem Speicher: Speicherslot dicke nehmen ; von einer Station die Scheibendicke nehmen
      *)
      IF ( starrShuttleBasisParameter[wStation].pAuftrag[wWand].rAuftragsDicke <= wgMKScheibenDicke13mm ) THEN
        starrShuttleBasisParameter[wStation].pAuftrag[wWand].stAuftragsOptionen.eDickenverstellung    := eZylinderStellung16mm;
      ELSIF ( starrShuttleBasisParameter[wStation].pAuftrag[wWand].rAuftragsDicke <= wgMKScheibenDicke19mm ) THEN
        starrShuttleBasisParameter[wStation].pAuftrag[wWand].stAuftragsOptionen.eDickenverstellung    := eZylinderStellung23mm;
      ELSIF ( starrShuttleBasisParameter[wStation].pAuftrag[wWand].rAuftragsDicke <= wgMKScheibenDicke24mm ) THEN
        starrShuttleBasisParameter[wStation].pAuftrag[wWand].stAuftragsOptionen.eDickenverstellung    := eZylinderStellung29mm;
      END_IF

      // Kippen
      starrShuttleBasisParameter[wStation].pAuftrag[wWand].stAuftragsOptionen.eKippen_SollPosition                  := starrShuttleBasisParameter[wStation].stMKs.stSchnittstellendaten.aEintransporte.Kippen[Auftragsdaten.wTransferstationsNr1];
      starrShuttleBasisParameter[wStation].pAuftrag[wWand].stAuftragsOptionen.eKippen_SollPosition_NachEintransport := starrShuttleBasisParameter[wStation].stMKs.stSchnittstellendaten.aEintransporte.KippenNachEintransport[Auftragsdaten.wTransferstationsNr1];
      starrShuttleBasisParameter[wStation].pAuftrag[wWand].stAuftragsOptionen.eKippen_SollPosition_NachAustransport := 0;

      // Hub
      starrShuttleBasisParameter[wStation].pAuftrag[wWand].stAuftragsOptionen.eHub                  := starrShuttleBasisParameter[wStation].stMKs.stSchnittstellendaten.aEintransporte.Hub[Auftragsdaten.wTransferstationsNr1];
      starrShuttleBasisParameter[wStation].pAuftrag[wWand].stAuftragsOptionen.eHub_NachEintransport := starrShuttleBasisParameter[wStation].stMKs.stSchnittstellendaten.aEintransporte.HubNachEintransport[Auftragsdaten.wTransferstationsNr1];
      starrShuttleBasisParameter[wStation].pAuftrag[wWand].stAuftragsOptionen.eHub_NachAustransport := 0;

      // Glastransport
      starrShuttleBasisParameter[wStation].pAuftrag[wWand].stAuftragsOptionen.eGlastransport := starrShuttleBasisParameter[wStation].stMKs.stSchnittstellendaten.aEintransporte.Glastransport[Auftragsdaten.wTransferstationsNr1];

      // Greifer [Ausbaustufe stStationsAufbau.bGreifer]: Greiferseite je Partnerstation, Zangenoeffnung wie die Scheibenfuehrung
      starrShuttleBasisParameter[wStation].pAuftrag[wWand].stAuftragsOptionen.eGreiferTyp := eGreiferDefault;
      IF ( starrShuttleBasisParameter[wStation].stMKs.stStationsAufbau.bGreifer[wWand] ) THEN
        starrShuttleBasisParameter[wStation].pAuftrag[wWand].stAuftragsOptionen.eGreiferTyp := starrShuttleBasisParameter[wStation].stMKs.stSchnittstellendaten.aEintransporte.Greifer[Auftragsdaten.wTransferstationsNr1];
      END_IF
      starrShuttleBasisParameter[wStation].pAuftrag[wWand].stAuftragsOptionen.eGreiferZangeStellung := starrShuttleBasisParameter[wStation].pAuftrag[wWand].stAuftragsOptionen.eDickenverstellung;

      // Scheibentyp prüfen
      starrShuttleBasisParameter[wStation].wGlasTyp[wWand] := eScheibe_Default;
      IF ( Auftragsdaten.rAuftragsLaenge >= starrShuttleBasisParameter[wStation].stMKs.stStationsParameter.rLaengeUebergroesseScheibe ) THEN
        starrShuttleBasisParameter[wStation].wGlasTyp[wWand] := eScheibe_Maximal;
      END_IF

      (* Anmerkung:
         - Zielstation abfragen ob diese bereit sind zum Austransport
           => Status der Glas-Sender Station pruefen
      *)
      CASE wlEintransportstation OF

        // Shuttles
        cERSTES_SHUTTLE..cLETZTES_SHUTTLE: // ... macht wenig Sinn
          ;

        // Transfershuttles
        cERSTES_TRANSFERSHUTTLE..cLETZTES_TRANSFERSHUTTLE:
          steplSchritt := STEP_200_E;

        // Stationen
        cERSTE_STATION..cLETZTE_STATION:
          IF ( ( Job_Stationen.AuftragsdatenWand[wlEintransportstation, Auftragsdaten.wTransferwand].wAuftrag = eStation_Warte_Auf_Austransport )
               OR ( Job_Stationen.AuftragsdatenWand[wlEintransportstation, Auftragsdaten.wTransferwand].wAuftrag = eStation_Belegt ) )
          THEN
            steplSchritt := STEP_100_E;
          END_IF

        cERSTE_FREMDANLAGE_AUSLAUF..cLETZTE_FREMDANLAGE_AUSLAUF:
          ;

        cERSTE_FREMDANLAGE_EINLAUF..cLETZTE_FREMDANLAGE_EINLAUF:
          ;

        // Faecherwagen direkt (Transferstation 1): nur mit dem Greifer. Ohne Greifer geht es aus dem Faecherwagen ueber ein
        // Transfershuttle mit bTransferShuttleFuerFaecherwagen (Transferstation 1 = Transfershuttle, Transferstation 2 = Faecherwagen)
        cERSTE_FAECHERWAGENSTATIONS_NR..cLETZTE_FAECHERWAGENSTATIONS_NR:
          IF ( starrShuttleBasisParameter[wStation].pAuftrag[wWand].stAuftragsOptionen.eGreiferTyp <> eGreiferDefault ) THEN
            IF ( starrFaecherwagenBasisParameter[wlEintransportstation].OutGlasTransport[cWAND_1].bBereitZumAustransport ) THEN
              steplSchritt := STEP_100_E;
            END_IF
          ELSE
            wpgFehlerdaten[0] := starrShuttleBasisParameter[wStation].stMKs.stStationsNummern.NummerExtern;
            wpgFehlerdaten[1] := wlEintransportstation;
            SpsError( eFehler_Station,
                      cMELDUNG_AUFTRAGSDATEN_FALSCHE_EINLAUFSTATION,
                      starrShuttleBasisParameter[wStation].stMKs.stStationsNummern.NummerIntern,
                      AutomatikkreisBestimmen(wStation),
                      wpgFehlerdaten );

            steplSchritt := STEP_900_E;
          END_IF

        ELSE
          wpgFehlerdaten[0] := starrShuttleBasisParameter[wStation].stMKs.stStationsNummern.NummerExtern;
          wpgFehlerdaten[1] := wlEintransportstation;
          SpsError( eFehler_Station,
                    cMELDUNG_AUFTRAGSDATEN_FALSCHE_EINLAUFSTATION,
                    starrShuttleBasisParameter[wStation].stMKs.stStationsNummern.NummerIntern,
                    AutomatikkreisBestimmen(wStation),
                    wpgFehlerdaten );

          steplSchritt := STEP_900_E;

      END_CASE

    // EINTRANSPORT ==============================================
    STEP_100_E:
      // ---------------------------------------------------------------------------------------
      //  EINTRANSPORT MITTELS STATIONEN [RKT, SF, ETC.]
      //
      //  Hinweis:
      // - n/c
      // ---------------------------------------------------------------------------------------

      (* Anmerkung:
         - Starten des Eintransports [Glas-Empfaenger]
         - Initiieren des  des Austransports [Glas-Empfaenger]
      *)
      CASE wlEintransportstation OF

        cERSTE_STATION..cLETZTE_STATION:

          IF AutomatikAktiv(wlEintransportstation) THEN

            (* Hinweis:
               - Auftragsdaten in Transferstation kopieren
            *)
            Job_Stationen.AuftragsdatenWand[wlEintransportstation, Auftragsdaten.wTransferwand]           := AuftragsdatenUmkopieren(FALSE, FALSE, Auftragsdaten);
            Job_Stationen.AuftragsdatenWand[wlEintransportstation, Auftragsdaten.wTransferwand].wAuftrag  := eStation_Austransport;

            (* Hinweis:
               - Kopplung zur Transferstation herstellen
            *)
            starrShuttleBasisParameter[wStation].InGlasTransportVorgaenger[wWand] := starrStationBasisParameter[wlEintransportstation].OutGlasTransport[Auftragsdaten.wTransferwand];
            starrShuttleBasisParameter[wStation].InGlasTransportNachfolger[wWand] := starrStationBasisParameter[wlEintransportstation].OutGlasTransport[Auftragsdaten.wTransferwand];

            (* Hinweis:
               - Starten des Eintransports
            *)
            starrShuttleBasisParameter[wStation].bScheibentrennen[wWand] := NOT Auftragsdaten.stAuftragsInformationen.cBIT_SRC_WALL_1_EMPTY;
            starrShuttleBasisParameter[wStation].bRueckwaertsTransportieren[wWand] := ( starrShuttleBasisParameter[wStation].stMKs.stSchnittstellendaten.aEintransporte.Station[wlEintransportstation] = Rueckwaertig );
            starrShuttleBasisParameter[wStation].bEintransport[wWand] := TRUE;

            steplSchritt := STEP_400_E;

          END_IF

        cERSTE_FREMDANLAGE_AUSLAUF..cLETZTE_FREMDANLAGE_AUSLAUF:
          ;

        cERSTE_FREMDANLAGE_EINLAUF..cLETZTE_FREMDANLAGE_EINLAUF:
          ;

        cERSTE_FAECHERWAGENSTATIONS_NR..cLETZTE_FAECHERWAGENSTATIONS_NR:
          (* Hinweis:
             - Eintransport aus dem Faecherwagen mit dem Greifer (Greiferseite im Auftrag)
          *)
          starrShuttleBasisParameter[wStation].bScheibentrennen[wWand]           := FALSE;
          starrShuttleBasisParameter[wStation].bRueckwaertsTransportieren[wWand] := FALSE;
          starrShuttleBasisParameter[wStation].bEintransport[wWand]              := TRUE;

          steplSchritt := STEP_400_E;

      END_CASE

    // EINTRANSPORT ==============================================
    STEP_200_E:
      // ---------------------------------------------------------------------------------------
      //  EINTRANSPORT MITTELS TRANSFERSHUTTLE
      //
      //  Hinweis:
      //  - Transferstation2 = 0   => Eintransport mit nur einem Transfershuttle
      //  - Transferstation2 <> 0  => Eintransport im Transfershuttle-Verbund
      // ---------------------------------------------------------------------------------------

      IF ( Auftragsdaten.wTransferstationsNr2 = 0 OR starrTransfershuttleBasisParameter[wlEintransportstation].stMKs.stStationsOptionen.stTransfershuttle.bTransferShuttleFuerFaecherwagen ) THEN

        IF (  ( Job_Shuttle.AuftragsdatenTransfershuttle[wlEintransportstation].wAuftrag = eStation_Kein_Auftrag ) ) THEN
          steplSchritt := STEP_210_E;
        END_IF

      ELSE
        VailiderenTransfershuttleVerbund ( wTransferstation1 := wlEintransportstation,
                                           wTransferstation2 := Auftragsdaten.wTransferstationsNr2 );

        IF (  ( Job_Shuttle.AuftragsdatenTransfershuttle[wlEintransportstation].wAuftrag = eStation_Kein_Auftrag )
             AND ( Job_Shuttle.AuftragsdatenTransfershuttle[Auftragsdaten.wTransferstationsNr2].wAuftrag  = eStation_Kein_Auftrag ) )
        THEN
          steplSchritt := STEP_220_E;
        END_IF

      END_IF

    // EINTRANSPORT ==============================================
    STEP_210_E:
      // ---------------------------------------------------------------------------------------
      //  EINTRANSPORT TRANSFERSHUTTLE [DEFAULT]
      //
      //  Hinweis:
      // - n/c
      // ---------------------------------------------------------------------------------------

      (* Hinweis:
         - Kopplung
      *)
      IF ( starrShuttleBasisParameter[wStation].stMKs.stSchnittstellendaten.aEintransporte.Station[wlEintransportstation] = Rueckwaertig ) THEN
        starrTransfershuttleBasisParameter[wlEintransportstation].InGlasTransportVorgaenger[wWand] := starrShuttleBasisParameter[wStation].OutGlasTransport[wWand];
        starrShuttleBasisParameter[wStation].InGlasTransportNachfolger[wWand] := starrTransfershuttleBasisParameter[wlEintransportstation].OutGlasTransport[wWand];

      ELSE
        starrTransfershuttleBasisParameter[wlEintransportstation].InGlasTransportNachfolger[wWand] := starrShuttleBasisParameter[wStation].OutGlasTransport[wWand];
        starrShuttleBasisParameter[wStation].InGlasTransportVorgaenger[wWand] := starrTransfershuttleBasisParameter[wlEintransportstation].OutGlasTransport[wWand];

      END_IF

      (* Hinweis:
         - TS auf FW koppeln
      *)
      IF   starrTransfershuttleBasisParameter[wlEintransportstation].stMKs.stStationsOptionen.stTransfershuttle.bTransferShuttleFuerFaecherwagen
           AND IsBetweenWORD(Auftragsdaten.wTransferstationsNr2, cERSTE_FAECHERWAGENSTATIONS_NR, cLETZTE_FAECHERWAGENSTATIONS_NR)
      THEN
        IF ( starrShuttleBasisParameter[wStation].stMKs.stSchnittstellendaten.aEintransporte.Station[wlEintransportstation] = Rueckwaertig ) THEN
          starrTransfershuttleBasisParameter[wlEintransportstation].InGlasTransportNachfolger[wWand] := starrFaecherwagenBasisParameter[Auftragsdaten.wTransferstationsNr2].OutGlasTransport[cWAND_1];
        ELSE
          starrTransfershuttleBasisParameter[wlEintransportstation].InGlasTransportVorgaenger[wWand] := starrFaecherwagenBasisParameter[Auftragsdaten.wTransferstationsNr2].OutGlasTransport[cWAND_1];
        END_IF
      END_IF

      (* Hinweis:
         - Neuen Auftag in den FIFO [Warteschlange] eintragen
      *)
      Job_Shuttle.AuftragsdatenTransfershuttle[wlEintransportstation]          := AuftragsdatenUmkopieren(FALSE, FALSE, Auftragsdaten);
      Job_Shuttle.AuftragsdatenTransfershuttle[wlEintransportstation].wAuftrag := eStation_Austransport;

      starrShuttleBasisParameter[wStation].bScheibentrennen[wWand]                := FALSE;
      starrShuttleBasisParameter[wStation].bRueckwaertsTransportieren[wWand]      := ( starrShuttleBasisParameter[wStation].stMKs.stSchnittstellendaten.aEintransporte.Station[wlEintransportstation] = Rueckwaertig );
      starrShuttleBasisParameter[wStation].bEintransport[wWand]                   := TRUE;
      starrShuttleBasisParameter[wStation].bTransferstationTransfershuttle[wWand] := TRUE;

      steplSchritt := STEP_400_E;

    // EINTRANSPORT ==============================================
    STEP_220_E:
      // ---------------------------------------------------------------------------------------
      //  EINTRANSPORT TRANSFERSHUTTLE [VERBUND]
      //
      //  Hinweis:
      //  - n/c
      // ---------------------------------------------------------------------------------------

      (* Hinweis:
         - Kopplung
      *)
      IF ( starrShuttleBasisParameter[wStation].stMKs.eStationsTyp = eInputshuttle ) THEN
        starrTransfershuttleBasisParameter[wlEintransportstation].InGlasTransportVorgaenger[cWAND_1] := starrShuttleBasisParameter[wStation].OutGlasTransport[wWand];
        starrShuttleBasisParameter[wStation].InGlasTransportNachfolger[wWand] := starrTransfershuttleBasisParameter[wlEintransportstation].OutGlasTransport[cWAND_1];

      ELSE
        starrTransfershuttleBasisParameter[wlEintransportstation].InGlasTransportNachfolger[cWAND_1] := starrShuttleBasisParameter[wStation].OutGlasTransport[wWand];
        starrShuttleBasisParameter[wStation].InGlasTransportVorgaenger[wWand] := starrTransfershuttleBasisParameter[wlEintransportstation].OutGlasTransport[cWAND_1];

      END_IF

      (* Hinweis:
         - Transfershuttle koppeln
      *)
      aTransfershuttles[wlEintransportstation].stpInTransportVerbund := aTransfershuttles[Auftragsdaten.wTransferstationsNr2].stpOutTransportVerbund;
      aTransfershuttles[Auftragsdaten.wTransferstationsNr2].stpInTransportVerbund  := aTransfershuttles[wlEintransportstation].stpOutTransportVerbund;

      (* Hinweis:
         - Auftragsdaten an die Transfershuttle uebergeben
      *)
      Job_Shuttle.AuftragsdatenTransfershuttle[wlEintransportstation]            := AuftragsdatenUmkopieren(FALSE, FALSE, Auftragsdaten);
      Job_Shuttle.AuftragsdatenTransfershuttle[wlEintransportstation].wAuftrag   := eStation_Austransport;

      Job_Shuttle.AuftragsdatenTransfershuttle[Auftragsdaten.wTransferstationsNr2]          := AuftragsdatenUmkopieren(TRUE, FALSE, Auftragsdaten);
      Job_Shuttle.AuftragsdatenTransfershuttle[Auftragsdaten.wTransferstationsNr2].wAuftrag := eStation_Transportkopplung;

      starrShuttleBasisParameter[wStation].bScheibentrennen[wWand]                := FALSE;
      starrShuttleBasisParameter[wStation].bRueckwaertsTransportieren[wWand]      := ( starrShuttleBasisParameter[wStation].stMKs.stSchnittstellendaten.aEintransporte.Station[wlEintransportstation] = Rueckwaertig );
      starrShuttleBasisParameter[wStation].bEintransport[wWand]                   := TRUE;
      starrShuttleBasisParameter[wStation].bTransferstationTransfershuttle[wWand] := TRUE;

      steplSchritt := STEP_400_E;

    // EINTRANSPORT ==============================================
    STEP_400_E:
      (* Hinweis:
         - Scheibenquittieren [pro Wand] -> Nachricht an die Oberflaeche
           =>( Oberflaeche prueft nicht die Wandnr. die quittiert werden nur bei einem multiplen  Ein-/Austransport- Auftrag wird die WandNr. geprueft )
      *)
      blStationQuittiertScheiben := starrShuttleBasisParameter[wStation].stMKs.stSchnittstellendaten.aEintransporte.bStationQuittiertScheibe[wlEintransportstation];

      IF ( starrShuttleBasisParameter[wStation].OutGlasTransport[wWand].bQuittScheibe ) THEN

        IF ( ilScheibenZuQuittieren > 0 ) AND blStationQuittiertScheiben THEN

          wSps2MmiZielStation  := starrShuttleBasisParameter[wStation].stMKs.stStationsNummern.NummerIntern;
          wSps2MmiQuellStation := Auftragsdaten.wTransferstationsNr1;
          wSps2MmiZielWand     := wWand;
          wSps2MmiQuellWand    := Auftragsdaten.wTransferwand;
          dwSps2MmiWartezeit   := starrShuttleBasisParameter[wStation].dwWartezeit[wWand];
          wSPS2MMIAuftragstyp  := 0;

          MsgToMmi(auftragsnr_w := SB0_SPS_QUIT_SHEET_ORDER );
        END_IF

        ilScheibenZuQuittieren := ilScheibenZuQuittieren - 1;

      END_IF

      (* Anmerkung:
         - Transport abgeschlossen
      *)
      IF ( starrShuttleBasisParameter[wStation].bEintransportAbgeschlossen[wWand] ) THEN
        starrShuttleBasisParameter[wStation].bEintransport[wWand] := FALSE;
        starrShuttleBasisParameter[wStation].bRueckwaertsTransportieren[wWand] := FALSE;
        steplSchritt := STEP_410_E;
      END_IF

      (* Fehlerbehandlung:
         - Shuttle
      *)
      IF ( starrShuttleBasisParameter[wStation].bFehler ) THEN
        SpsError( eFehler_Station,
                  starrShuttleBasisParameter[wStation].wFehlerNummer,
                  starrShuttleBasisParameter[wStation].stMKs.stStationsNummern.NummerIntern,
                  AutomatikkreisBestimmen(wStation),
                  starrShuttleBasisParameter[wStation].awFehlerInformationen );

        starrShuttleBasisParameter[wStation].bEintransport[wWand] := FALSE;
        starrShuttleBasisParameter[wStation].bRueckwaertsTransportieren[wWand] := FALSE;

        steplSchritt := STEP_900_E;

      END_IF

    // EINTRANSPORT ==============================================
    STEP_410_E:
      (* Anmerkung:
         - Gueltige Anzahl von Scheiben wurden quittiert
      *)
      IF ( ilScheibenZuQuittieren = 0 ) THEN

        steplSchritt := STEP_1000_E;

      (* Anmerkung:
         - Zu wenig Scheiben quittiert
      *)
      ELSIF ( ilScheibenZuQuittieren > 0 ) THEN
        wpgFehlerdaten[0] := starrShuttleBasisParameter[wStation].stMKs.stStationsNummern.NummerExtern;
        wpgFehlerdaten[1] := wWand;

        SpsError( eFehler_Station,
                  cMELDUNG_STATION_ZUWENIG_SCHEIBEN_QUITTIERT_WAND_EINTRANSPORT,
                  starrShuttleBasisParameter[wStation].stMKs.stStationsNummern.NummerIntern,
                  AutomatikkreisBestimmen(wStation),
                  wpgFehlerdaten );

        steplSchritt := STEP_900_E;

      (* Anmerkung:
         - Zu viele Scheiben quittiert
      *)
      ELSIF ( ilScheibenZuQuittieren < 0 )  THEN
        wpgFehlerdaten[0] := starrShuttleBasisParameter[wStation].stMKs.stStationsNummern.NummerExtern;
        wpgFehlerdaten[1] := wWand;

        SpsError( eFehler_Station,
                  cMELDUNG_STATION_ZUVIELE_SCHEIBEN_QUITTIERT_WAND_EINTRANSPORT,
                  starrShuttleBasisParameter[wStation].stMKs.stStationsNummern.NummerIntern,
                  AutomatikkreisBestimmen(wStation),
                  wpgFehlerdaten );

        steplSchritt := STEP_900_E;

      END_IF

    // EINTRANSPORT ==============================================
    STEP_900_E:
      starrShuttleBasisParameter[wStation].bEintransport[wWand] := FALSE;
      starrShuttleBasisParameter[wStation].bRueckwaertsTransportieren[wWand] := FALSE;

      bpFehler := TRUE;

    // EINTRANSPORT ==============================================
    STEP_1000_E:
      (* Hinweis:
         - Beenden des Eintransports [Bereit fuer den naechsten Auftrag]
      *)
      bpDone := TRUE;
      Auftragsdaten.wAuftrag := eStation_Kein_Auftrag;

  // EINTRANSPORT ==============================================
  END_CASE
END_IF

IF bpReset THEN
  bpFehler := FALSE;
  bpDone := FALSE;
  bpReset := FALSE;
  starrShuttleBasisParameter[wStation].bEintransport[wWand] := FALSE;
  starrShuttleBasisParameter[wStation].bRueckwaertsTransportieren[wWand] := FALSE;
  starrShuttleBasisParameter[wStation].bTransferstationTransfershuttle[wWand] := FALSE;
  steplSchritt := STEP_0_E;
END_IF
END_FUNCTION_BLOCK

(* ---- Shuttle_Querfahrt.fb.st ---- *)
(* METADATA
{
	"v3Meta": {
		"objectGuid": "b8d8b63a-039c-49d7-ab0c-8520bb128b08"
	}
}
*)
FUNCTION_BLOCK Shuttle_Querfahrt
VAR_INPUT

  // BOOLEAN
  bpReset                : BOOL;

  // WORD
  wStation               : WORD;

  // STRUKTUR
  Auftragsdaten          : Auftragsdaten_ST;

END_VAR
VAR_OUTPUT

  // BOOL
  bpDone                 : BOOL;
  bpFehler               : BOOL;

END_VAR
VAR

  // STEPS
  steplSchritt                    : STEPS_TE;

  // BAUSTEINE
  PositionierAuftragsdatenPruefen : PositionierAuftragsdatenPruefen;

END_VAR
// ****************************************************9*********************************************
// STEUERUNG: POSITIONIEREN
// *************************************************************************************************

IF ( Auftragsdaten.wAuftrag = eStation_Vorabpositionierung ) THEN
  CASE steplSchritt OF
    // POSITIONIERUNG ===========================================
    STEP_0_E:
      (* Hinweis:
         - Ueberpruefung des Sicherheitskreises
      *)
      IF checkSafetyCircuitsNotBlocked(starrShuttleBasisParameter[wStation]) THEN

        IF ( ABS( starrShuttleBasisParameter[wStation].rAktuellePositionQuerfahrt - Auftragsdaten.rVorabPosition ) <= rgMKZielPositionToleranz ) THEN
          steplSchritt := STEP_500_E;
        ELSIF starrShuttleBasisParameter[wStation].stMKs.bDeaktivieren THEN
          steplSchritt := STEP_600_E;
        ELSE
          steplSchritt := STEP_5_E;
        END_IF

      END_IF

    // POSITIONIERUNG ===========================================
    STEP_5_E:
      (* Hinweis:
         - Auftragsdaten pruefen
           => Version der Verfahrlogik beachten
      *)
      steplSchritt := STEP_10_E;

      PositionierAuftragsdatenPruefen.rpSollPosition   := Auftragsdaten.rVorabPosition;
      PositionierAuftragsdatenPruefen.wpStationsNummer := wStation;

      PositionierAuftragsdatenPruefen();

      IF ( NOT PositionierAuftragsdatenPruefen.bpErgebnis ) THEN
        steplSchritt := STEP_900_E;
      END_IF

    // POSITIONIERUNG ===========================================
    STEP_10_E:
      (* Hinweis:
         - Uebergabe der Auftragsdaten
      *)
      starrShuttleBasisParameter[wStation].pAuftragVorabPositionierung := Auftragsdaten;
      starrShuttleBasisParameter[wStation].bVorabpositionieren := TRUE;

      steplSchritt := STEP_20_E;

    // POSITIONIERUNG ===========================================
    STEP_20_E:
      (* Hinweis:
         - Nachricht absetzen
      *)
      IF ( starrShuttleBasisParameter[wStation].bUpdateVorabPositionieren = TRUE ) THEN

        wSps2MmiQuittVorabShuttleNr := starrShuttleBasisParameter[wStation].stMKs.stStationsNummern.NummerIntern;
        rgSPS2MMIExtractionShuttlePosition := starrShuttleBasisParameter[wStation].rAktuellePositionQuerfahrt;
        MsgToMmi(auftragsnr_w := SB0_SPS_SHUTTLEVORABPOSITIONIERUNGUPDATE );// Quit 2 MMI Scheibe vorne

        starrShuttleBasisParameter[wStation].bUpdateVorabPositionieren := FALSE;

        steplSchritt := STEP_100_E;

      END_IF

      (* Fehlerbehandlung:
         - Inputshuttle
      *)
      IF ( starrShuttleBasisParameter[wStation].bFehler ) THEN

        starrShuttleBasisParameter[wStation].bVorabpositionieren := FALSE;

        SpsError( eFehler_Station,
                  starrShuttleBasisParameter[wStation].wFehlerNummer,
                  starrShuttleBasisParameter[wStation].stMKs.stStationsNummern.NummerIntern,
                  AutomatikkreisBestimmen(starrShuttleBasisParameter[wStation].stMKs.stStationsNummern.NummerSPS),
                  starrShuttleBasisParameter[wStation].awFehlerInformationen );

        steplSchritt := STEP_900_E;
      END_IF

    // POSITIONIERUNG ===========================================
    STEP_100_E:
      (* Hinweis:
         - Positionierung abgeschlossen
           => Nachricht absetzen
      *)
      IF ( starrShuttleBasisParameter[wStation].bVorabpositionierenAbgeschlossen ) THEN

        starrShuttleBasisParameter[wStation].bVorabpositionieren := FALSE;

        wSps2MmiQuittVorabShuttleNr        := starrShuttleBasisParameter[wStation].stMKs.stStationsNummern.NummerIntern;
        rgSPS2MMIExtractionShuttlePosition := starrShuttleBasisParameter[wStation].rAktuellePositionQuerfahrt;
        MsgToMmi(auftragsnr_w := SB0_SPS_QUITTSHUTTLEVORABPOSITIONIERUNG );

        steplSchritt := STEP_1000_E;

      END_IF

      (* Fehlerbehandlung:
         - Inputshuttle
      *)
      IF ( starrShuttleBasisParameter[wStation].bFehler ) THEN
        starrShuttleBasisParameter[wStation].bVorabpositionieren := FALSE;

        SpsError( eFehler_Station,
                  starrShuttleBasisParameter[wStation].wFehlerNummer,
                  starrShuttleBasisParameter[wStation].stMKs.stStationsNummern.NummerIntern,
                  AutomatikkreisBestimmen(starrShuttleBasisParameter[wStation].stMKs.stStationsNummern.NummerSPS),
                  starrShuttleBasisParameter[wStation].awFehlerInformationen );

        steplSchritt := STEP_900_E;
      END_IF

    // POSITIONIERUNG ===========================================
    STEP_500_E:
      wSps2MmiQuittVorabShuttleNr := starrShuttleBasisParameter[wStation].stMKs.stStationsNummern.NummerIntern;
      rgSPS2MMIExtractionShuttlePosition := starrShuttleBasisParameter[wStation].rAktuellePositionQuerfahrt;
      MsgToMmi(auftragsnr_w := SB0_SPS_SHUTTLEVORABPOSITIONIERUNGUPDATE );
      steplSchritt := STEP_510_E;

    // POSITIONIERUNG ===========================================
    STEP_510_E:
      wSps2MmiQuittVorabShuttleNr        := starrShuttleBasisParameter[wStation].stMKs.stStationsNummern.NummerIntern;
      rgSPS2MMIExtractionShuttlePosition := starrShuttleBasisParameter[wStation].rAktuellePositionQuerfahrt;
      MsgToMmi(auftragsnr_w := SB0_SPS_QUITTSHUTTLEVORABPOSITIONIERUNG );
      steplSchritt := STEP_1000_E;

    // POSITIONIERUNG ===========================================
    STEP_600_E:
      wSps2MmiQuittVorabShuttleNr := starrShuttleBasisParameter[wStation].stMKs.stStationsNummern.NummerIntern;
      rgSPS2MMIExtractionShuttlePosition := Auftragsdaten.rVorabPosition;
      MsgToMmi(auftragsnr_w := SB0_SPS_SHUTTLEVORABPOSITIONIERUNGUPDATE );
      steplSchritt := STEP_610_E;

    // POSITIONIERUNG ===========================================
    STEP_610_E:
      wSps2MmiQuittVorabShuttleNr        := starrShuttleBasisParameter[wStation].stMKs.stStationsNummern.NummerIntern;
      rgSPS2MMIExtractionShuttlePosition := Auftragsdaten.rVorabPosition;
      MsgToMmi(auftragsnr_w := SB0_SPS_QUITTSHUTTLEVORABPOSITIONIERUNG );
      steplSchritt := STEP_1000_E;

    // POSITIONIERUNG ===========================================
    STEP_900_E:
      bpFehler := TRUE;

    // POSITIONIERUNG ===========================================
    STEP_1000_E:
      bpDone := TRUE;
      Auftragsdaten.wAuftrag := eStation_Kein_Auftrag;

  // POSITIONIERUNG ===========================================
  END_CASE
END_IF

IF bpReset THEN
  bpFehler := FALSE;
  bpDone := FALSE;
  bpReset := FALSE;
  starrShuttleBasisParameter[wStation].bUpdateVorabPositionieren := FALSE;
  starrShuttleBasisParameter[wStation].bVorabpositionieren := FALSE;
  steplSchritt := STEP_0_E;
END_IF
END_FUNCTION_BLOCK

(* ---- Shuttle_RackSuche.fb.st ---- *)
(* METADATA
{
	"v3Meta": {
		"objectGuid": "f075b551-e071-4bf5-ac95-2cac71043e2d"
	}
}
*)
FUNCTION_BLOCK Shuttle_RackSuche
VAR_INPUT

  // BOOLEAN
  bpReset                : BOOL;

  // WORD
  wStation               : WORD;

  // STRUKTUR
  Auftragsdaten          : Auftragsdaten_ST;

END_VAR
VAR_OUTPUT

  // BOOLEAN
  bpDone                 : BOOL;
  bpFehler               : BOOL;

END_VAR
VAR

  // STEPS
  steplSchritt           : STEPS_TE;

END_VAR
//-------------------------------------------------------------------------------------------------
// STEUERUNG VORABKOMPONENETEN
//-------------------------------------------------------------------------------------------------

IF ( Auftragsdaten.wAuftrag = eStation_RackSuche ) THEN

  (* Fehlerbehandlung:
     - Inputshuttle
  *)
  IF starrShuttleBasisParameter[wStation].bFehler AND steplSchritt <> STEP_900_E THEN
    aShuttle[wStation].bpStarteFaecherwagensuche := FALSE;
    SpsError( eFehler_Station,
              starrShuttleBasisParameter[wStation].wFehlerNummer,
              starrShuttleBasisParameter[wStation].stMKs.stStationsNummern.NummerIntern,
              AutomatikkreisBestimmen(wStation),
              starrShuttleBasisParameter[wStation].awFehlerInformationen );

    steplSchritt := STEP_900_E;
  END_IF

  CASE steplSchritt OF
    // RACKSUCHE ===========================================
    STEP_0_E:
      (* Hinweis:
         - Pruefen ob der Sicherheitskreis ausgeloest oder angefragz wurde
      *)
      IF checkSafetyCircuitsNotBlocked(starrShuttleBasisParameter[wStation]) THEN
        steplSchritt := STEP_10_E;
      END_IF

    // RACKSUCHE ===========================================
    STEP_10_E:
      (* Hinweis:
         - Starten der Schrittkette -> MMI Fährt mittel Shuttlepositionierung den Weg ab
      *)
      aShuttle[wStation].bpStarteFaecherwagensuche := TRUE;

      steplSchritt := STEP_100_E;

    // RACKSUCHE ===========================================
    STEP_100_E:
      (* Hinweis:
         - Fächerwagensuche: Wort 0 = (int) SPS Nr Shuttle  / Wort 1+2 = (real) Position rechte (?) Kante der Folie[-1 für nicht gefunden]
           => Nachricht absetzen
      *)
      IF ( aShuttle[wStation].bpFaecherwagenGefunden ) THEN

        wSps2MmiStationsNummer     := starrShuttleBasisParameter[wStation].stMKs.stStationsNummern.NummerIntern;
        rSps2MmiPosition           := aShuttle[wStation].rpAktuelleFaecherwagenPosition;
        MsgToMmi(auftragsnr_w := SB0_SPS_POSITIONMEASUREDATA );

        steplSchritt := STEP_1000_E;

      END_IF

    // RACKSUCHE ===========================================
    STEP_900_E:
      bpFehler := TRUE;

    // RACKSUCHE ===========================================
    STEP_1000_E:
      bpDone := TRUE;
      Auftragsdaten.wAuftrag := eStation_Kein_Auftrag;

  // RACKSUCHE ===========================================
  END_CASE

END_IF

IF bpReset THEN
  bpFehler := FALSE;
  bpDone := FALSE;
  bpReset := FALSE;
  aShuttle[wStation].bpStarteFaecherwagensuche := FALSE;
  IF (aShuttle[wStation].rpAktuelleFaecherwagenPosition = -100000)  THEN // ungültige Rackposition von -10000 angeben da kein Rack gefunden
    wSps2MmiStationsNummer     := starrShuttleBasisParameter[wStation].stMKs.stStationsNummern.NummerIntern;
    rSps2MmiPosition           := aShuttle[wStation].rpAktuelleFaecherwagenPosition;
    MsgToMmi(auftragsnr_w := SB0_SPS_POSITIONMEASUREDATA );
  END_IF
  steplSchritt := STEP_0_E;
END_IF
END_FUNCTION_BLOCK

(* ---- Shuttle_Vorabkomponenten.fb.st ---- *)
(* METADATA
{
	"v3Meta": {
		"objectGuid": "19fcb8bb-2bd9-4575-a4db-49bc1e849a70"
	}
}
*)
FUNCTION_BLOCK Shuttle_Vorabkomponenten
VAR_INPUT

  // BOOLEAN
  bpReset                : BOOL;

  // WORD
  wStation               : WORD;
  wWand                  : WORD;

  // STRUKTUR
  Auftragsdaten          : VorAbAuftragsdaten_ST;

END_VAR
VAR_OUTPUT

  // BOOLEAN
  bpDone                 : BOOL;
  bpFehler               : BOOL;

END_VAR
VAR

  // BOOL
  blFreigabeVorabAuftrag     : BOOL;

  // WORD
  wlNextTransferstation  : WORD;

  // STEPS
  steplSchritt           : STEPS_TE;

END_VAR
//-------------------------------------------------------------------------------------------------
// STEUERUNG VORABKOMPONENETEN
//-------------------------------------------------------------------------------------------------

IF ( Auftragsdaten.wAuftrag = eStation_VorabAuftrag ) THEN

  (* Hinweis:
     - Setzen der Freigabe fuer die Resourcen-Ansteuerung wenn zum Zeitpunkt des "STARTENS"
       kein Auftrag aktiv ist. Ist die Ansteuerung "Aktiv" kann diese Variable wieder abfallen.
  *)
  blFreigabeVorabAuftrag := ( Job_Shuttle.AuftragsdatenWand[wStation, wWand].wAuftrag = eStation_Kein_Auftrag );

  CASE steplSchritt OF

    // VORABKOMPONENETEN ===============================================
    STEP_0_E:
      (* Hinweis:
         - Ueberpruefung des Sicherheitskreises
      *)
      IF checkSafetyCircuitsNotBlocked(starrShuttleBasisParameter[wStation])
         AND blFreigabeVorabAuftrag
      THEN
        IF ( Auftragsdaten.wTransferStation <> 0 ) THEN
          steplSchritt := STEP_10_E;
        ELSE
          steplSchritt := STEP_1000_E;
        END_IF
      END_IF

    // VORABKOMPONENETEN ===============================================
    STEP_10_E:
      // Transferstation bestimmen
      wlNextTransferstation := Auftragsdaten.wTransferStation;

      // Auftragsdaten uebergeben
      starrShuttleBasisParameter[wStation].pVorAbAuftragsdaten[wWand]:= Auftragsdaten;

      // Vorinitialisieren der Werte
      starrShuttleBasisParameter[wStation].pVorAbAuftragsdaten[wWand].stAuftragsOptionen.eGlastransport       := eGlastransport_Default;
      starrShuttleBasisParameter[wStation].pVorAbAuftragsdaten[wWand].stAuftragsOptionen.eDickenverstellung   := eZylinderUndefiniert;
      starrShuttleBasisParameter[wStation].pVorAbAuftragsdaten[wWand].stAuftragsOptionen.eKippen_SollPosition := eKippen_Default;

      // Scheibentyp prüfen
      starrShuttleBasisParameter[wStation].wGlasTyp[wWand] := eScheibe_Default;
      IF ( Auftragsdaten.rLaenge >= starrShuttleBasisParameter[wStation].stMKs.stStationsParameter.rLaengeUebergroesseScheibe ) THEN
        starrShuttleBasisParameter[wStation].wGlasTyp[wWand] := eScheibe_Maximal;
      END_IF

      (* Hinweis:
         - Austransport
      *)
      IF ( Auftragsdaten.wAuftragstyp.0 ) THEN
        // Folgestation beruecksichtigen damit in verschiedene Richtungen vorpositioniert werden kann.
        starrShuttleBasisParameter[wStation].pVorAbAuftragsdaten[wWand].stAuftragsOptionen.eGlastransport := starrShuttleBasisParameter[wStation].stMKs.stSchnittstellendaten.aAustransporte.Glastransport[wlNextTransferstation];
        starrShuttleBasisParameter[wStation].pVorAbAuftragsdaten[wWand].stAuftragsOptionen.eKippen_SollPosition := starrShuttleBasisParameter[wStation].stMKs.stSchnittstellendaten.aAustransporte.Kippen[wlNextTransferstation];
      ELSE
        starrShuttleBasisParameter[wStation].pVorAbAuftragsdaten[wWand].stAuftragsOptionen.eKippen_SollPosition := starrShuttleBasisParameter[wStation].stMKs.stSchnittstellendaten.aEintransporte.Kippen[wlNextTransferstation];
      END_IF

      // Greifer [Ausbaustufe stStationsAufbau.bGreifer]: Greiferseite je Partnerstation fuer die Vorabpositionierung
      starrShuttleBasisParameter[wStation].pVorAbAuftragsdaten[wWand].stAuftragsOptionen.eGreiferTyp := eGreiferDefault;
      IF ( starrShuttleBasisParameter[wStation].stMKs.stStationsAufbau.bGreifer[wWand] ) THEN
        IF ( Auftragsdaten.wAuftragstyp.0 ) THEN
          starrShuttleBasisParameter[wStation].pVorAbAuftragsdaten[wWand].stAuftragsOptionen.eGreiferTyp := starrShuttleBasisParameter[wStation].stMKs.stSchnittstellendaten.aAustransporte.Greifer[wlNextTransferstation];
        ELSE
          starrShuttleBasisParameter[wStation].pVorAbAuftragsdaten[wWand].stAuftragsOptionen.eGreiferTyp := starrShuttleBasisParameter[wStation].stMKs.stSchnittstellendaten.aEintransporte.Greifer[wlNextTransferstation];
        END_IF
      END_IF

      (* Hinweis:
         - Scheibenführung / Wandverstellung anstellen
         - Aus dem Speicher: Speicherslotdicke nehmen ; von einer Station die Scheibendicke nehmen
      *)
      IF ( starrShuttleBasisParameter[wStation].pAuftrag[cWAND_1].rAuftragsDicke <= wgMKScheibenDicke13mm ) THEN
        starrShuttleBasisParameter[wStation].pVorAbAuftragsdaten[wWand].stAuftragsOptionen.eDickenverstellung := eZylinderStellung16mm;
      ELSIF ( starrShuttleBasisParameter[wStation].pAuftrag[cWAND_1].rAuftragsDicke <= wgMKScheibenDicke19mm ) THEN
        starrShuttleBasisParameter[wStation].pVorAbAuftragsdaten[wWand].stAuftragsOptionen.eDickenverstellung := eZylinderStellung23mm;
      ELSIF ( starrShuttleBasisParameter[wStation].pAuftrag[cWAND_1].rAuftragsDicke <= wgMKScheibenDicke24mm ) THEN
        starrShuttleBasisParameter[wStation].pVorAbAuftragsdaten[wWand].stAuftragsOptionen.eDickenverstellung := eZylinderStellung29mm;
      END_IF

      // Auftrag übergeben
      starrShuttleBasisParameter[wStation].bVorabKomponentenAnsteuerung[wWand] := TRUE;

      steplSchritt := STEP_400_E;

    // VORABKOMPONENETEN ===============================================
    STEP_400_E:
      (* Hinweis:
         - Abschliessen des Austransports
      *)
      IF ( starrShuttleBasisParameter[wStation].bVorabKomponentenAnsteuerungAbgeschlossen[wWand] ) THEN
        starrShuttleBasisParameter[wStation].bVorabKomponentenAnsteuerung[wWand] := FALSE;
        steplSchritt := STEP_1000_E;
      END_IF

      (* Fehlerbehandlung:
         - Inputshuttle
      *)
      IF ( starrShuttleBasisParameter[wStation].bFehler ) THEN
        SpsError( eFehler_Station,
                  starrShuttleBasisParameter[wStation].wFehlerNummer,
                  starrShuttleBasisParameter[wStation].stMKs.stStationsNummern.NummerIntern,
                  AutomatikkreisBestimmen(starrShuttleBasisParameter[wStation].stMKs.stStationsNummern.NummerSPS),
                  starrShuttleBasisParameter[wStation].awFehlerInformationen );

        steplSchritt := STEP_900_E;
      END_IF

    // VORABKOMPONENETEN ===============================================
    STEP_900_E:
      blFreigabeVorabAuftrag := FALSE;
      bpFehler := TRUE;

    // VORABKOMPONENETEN ===============================================
    STEP_1000_E:
      bpDone := TRUE;
      blFreigabeVorabAuftrag := FALSE;
      Auftragsdaten.wAuftrag := eStation_Kein_Auftrag;

  // VORABKOMPONENETEN ===============================================
  END_CASE

END_IF

IF bpReset THEN
  bpFehler := FALSE;
  bpDone := FALSE;
  bpReset := FALSE;
  blFreigabeVorabAuftrag := FALSE;
  starrShuttleBasisParameter[wStation].bVorabKomponentenAnsteuerung[wWand] := FALSE;
  steplSchritt := STEP_0_E;
END_IF
END_FUNCTION_BLOCK

(* ---- Station_Abnehmen.fb.st ---- *)
(* METADATA
{
	"v3Meta": {
		"objectGuid": "c33fea17-eb20-4bc7-9a81-45f784503e7d"
	}
}
*)
FUNCTION_BLOCK Station_Abnehmen
VAR_INPUT

  // BOOLEAN
  bpReset                : BOOL;

  // WORD
  wStation               : WORD;

  // STRUKTUR
  Auftragsdaten          : Auftragsdaten_ST;

END_VAR
VAR_OUTPUT

  // BOOLEAN
  bpDone                 : BOOL;
  bpFehler               : BOOL;

END_VAR
VAR

  // INT
  ilScheibenZuQuittieren :  INT;

  // STEPS
  steplSchritt           : STEPS_TE;

END_VAR

//-------------------------------------------------------------------------------------------------
// STEUERUNG ABNEHMEN
//-------------------------------------------------------------------------------------------------
IF ( Auftragsdaten.wAuftrag = eStation_Abnehmen ) THEN
  CASE steplSchritt OF
    // ABNEHMEN =================================
    STEP_0_E:
      (* Hinweis:
         - Ueberpruefung des Sicherheitskreises
      *)
      IF checkSafetyCircuitsNotBlocked(starrStationBasisParameter[wStation]) THEN
        steplSchritt := STEP_10_E;
      END_IF

    // ABNEHMEN =================================
    STEP_10_E:
      starrStationBasisParameter[wStation].pAuftrag[cWAND_1] := Auftragsdaten;
      starrStationBasisParameter[wStation].bAbnehmen := TRUE;

      steplSchritt := STEP_20_E;

    // ABNEHMEN =================================
    STEP_20_E:
      IF (  starrStationBasisParameter[wStation].OutGlasTransport[cWAND_1].bQuittScheibe
           AND ilScheibenZuQuittieren > 0 )
      THEN
        ilScheibenZuQuittieren := ilScheibenZuQuittieren - 1;
      END_IF

      IF (ilScheibenZuQuittieren <= 0 ) THEN
        steplSchritt := STEP_30_E;
      END_IF

    // ABNEHMEN =================================
    STEP_30_E:
      (* Hinweis:
         - Glas wurde abgenommen
      *)
      IF ( starrStationBasisParameter[wStation].bAbnehmenAbgeschlossen ) THEN
        starrStationBasisParameter[wStation].bAbnehmen := FALSE;

        // Nachricht:
        //   - Das der Bediener die Scheibe abgenommen hat
        //     => Quittierung fuer Glas abgenommen
        //   - Nachricht dient nur zur Ueberwachung
        //   Wichtig:
        //   - Es kann sich aber immer noch Glas auf der Station befinden wenn der Bediener die Scheibe nicht entfernt hat
        wSps2MmiStationsNummer := starrStationBasisParameter[wStation].stMKs.stStationsNummern.NummerIntern;
        MsgToMmi(auftragsnr_w := SB0_SPS_SHEETREMOVEDAPPROVALWALL);

        steplSchritt := STEP_1000_E;
      END_IF

      (* Fehlerbehandlung:
         - Anlegewand
      *)
      IF ( starrStationBasisParameter[wStation].bFehler ) THEN
        SpsError( eFehler_Station,
                  starrStationBasisParameter[wStation].wFehlerNummer,
                  starrStationBasisParameter[wStation].stMKs.stStationsNummern.NummerIntern,
                  AutomatikkreisBestimmen(starrStationBasisParameter[wStation].stMKs.stStationsNummern.NummerSPS),
                  starrStationBasisParameter[wStation].awFehlerInformationen );

        starrStationBasisParameter[wStation].bAbnehmen := FALSE;
        steplSchritt := STEP_900_E;
      END_IF

    // ABNEHMEN =================================
    STEP_900_E:
      bpFehler := TRUE;

    // ABNEHMEN =================================
    STEP_1000_E:
      bpDone := TRUE;
      Auftragsdaten.wAuftrag := eStation_Kein_Auftrag;

  // ABNEHMEN =================================
  END_CASE
END_IF

IF bpReset THEN
  bpFehler := FALSE;
  bpDone := FALSE;
  bpReset := FALSE;
  steplSchritt := STEP_0_E;
  starrStationBasisParameter[wStation].bAbnehmen := FALSE;
END_IF
END_FUNCTION_BLOCK

(* ---- Station_Anlegen.fb.st ---- *)
(* METADATA
{
	"v3Meta": {
		"objectGuid": "d4215ee0-47ee-45d9-8520-4f4f5fb6c469"
	}
}
*)
FUNCTION_BLOCK Station_Anlegen
VAR_INPUT

  // BOOLEAN
  bpReset                : BOOL;
  bpAbbruchAnlegeauftrag : BOOL;

  // WORD
  wStation               : WORD;

  // STRUKTUR
  Auftragsdaten          : Auftragsdaten_ST;

END_VAR
VAR_OUTPUT

  // BOOLEAN
  bpDone                 : BOOL;
  bpFehler               : BOOL;

END_VAR
VAR

  // BOOL
  blAktiv                : BOOL;

  // STEPS
  steplSchritt           : STEPS_TE;

END_VAR

blAktiv := TRUE;
//-------------------------------------------------------------------------------------------------
// STEUERUNG ANLEGEN
//-------------------------------------------------------------------------------------------------
IF ( Auftragsdaten.wAuftrag = eStation_Anlegen ) THEN
  CASE steplSchritt OF
    // ANLEGEN ==================================================
    STEP_0_E:
      (* Hinweis:
         - Ueberpruefung des Sicherheitskreises
      *)
      IF checkSafetyCircuitsNotBlocked(starrStationBasisParameter[wStation]) THEN
        steplSchritt := STEP_10_E;
      END_IF

      (* Hinweis:
         - Abbruch des Anl
      *)
      IF ( bpAbbruchAnlegeauftrag ) THEN
        bpAbbruchAnlegeauftrag := FALSE;
        bpDone := TRUE;
        Auftragsdaten.wAuftrag := eStation_Kein_Auftrag;
      END_IF

    // ANLEGEN ==================================================
    STEP_10_E:
      // ---------------------------------------------------------------------------------------
      //  PRUEFUNG DER GLASDATEN [AUFTRAGSDATEN]
      //
      //  Hinweis:
      // - Anlegeauftraege muessen immer auf richte GLas- Abmessungen geprueft werden
      // ---------------------------------------------------------------------------------------
      steplSchritt := STEP_20_E;

      IF NOT AuftragsdatenPruefen( wStation, cWAND_1, Auftragsdaten) THEN
        steplSchritt := STEP_900_E;
      END_IF

    // ANLEGEN ==================================================
    STEP_20_E:
      (* Hinweis:
         - Starten des Anlegevorgangs
      *)

      // Glastyp bestimmen
      IF Auftragsdaten.bModell THEN
        starrStationBasisParameter[wStation].wGlasTyp[cWAND_1] := cMODELLSCHEIBE;
      ELSE
        starrStationBasisParameter[wStation].wGlasTyp[cWAND_1] := cDEFAULTSCHEIBE;
      END_IF

      starrStationBasisParameter[wStation].pAuftrag[cWAND_1] := Auftragsdaten;
      starrStationBasisParameter[wStation].bAnlegen := TRUE;

      steplSchritt := STEP_30_E;

    // ANLEGEN ==================================================
    STEP_30_E:
      (* Hinweis:
         - Prüfen dass der Auftragsstatus sich geändert hat
      *)
      IF ( starrStationBasisParameter[wStation].eStatusAuftrag = eAuftragAktiv )
         OR  ( starrStationBasisParameter[wStation].eStatusAuftrag = eAuftragAktivWiederholen )
      THEN
        steplSchritt := STEP_100_E;
      END_IF

    // ANLEGEN ==================================================
    STEP_100_E:
      (* Hinweis:
         - Station hat ihren Vorgang abgeschlossen
      *)
      IF ( starrStationBasisParameter[wStation].bAnlegenAbgeschlossen ) THEN
        starrStationBasisParameter[wStation].bAnlegen := FALSE;

        IF ( starrStationBasisParameter[wStation].eStatusAuftrag = eAuftragErfolgreich ) THEN

          wSps2MmiInputtableNummer := starrStationBasisParameter[wStation].stMKs.stStationsNummern.NummerIntern;
          dwSps2MmiWartezeit       := starrStationBasisParameter[wStation].dwWartezeit[cWAND_1];
          MsgToMmi(auftragsnr_w := SB0_SPS_SHEETONINPUTTABLE);

          IF Auftragsdaten.bModell OR NOT (starrStationBasisParameter[wStation].stMKs.stStationsOptionen.stGlastransport.bScheibenVermessen) THEN
            wSps2MmiInputtableNummer := starrStationBasisParameter[wStation].stMKs.stStationsNummern.NummerIntern;
            dwSps2MmiWartezeit       := starrStationBasisParameter[wStation].dwWartezeit[cWAND_1];
            MsgToMmi(auftragsnr_w := SB0_SPS_SortierungQuittInputInQueue);
          END_IF

        END_IF

        steplSchritt := STEP_1000_E;
      END_IF

      (* Fehlerbehandlung:
         - Anlegewand
      *)
      IF ( starrStationBasisParameter[wStation].bFehler ) THEN

        SpsError( eFehler_Station,
                  starrStationBasisParameter[wStation].wFehlerNummer,
                  starrStationBasisParameter[wStation].stMKs.stStationsNummern.NummerIntern,
                  AutomatikkreisBestimmen(starrStationBasisParameter[wStation].stMKs.stStationsNummern.NummerSPS),
                  starrStationBasisParameter[wStation].awFehlerInformationen );

        starrStationBasisParameter[wStation].bAnlegen := FALSE;
        steplSchritt := STEP_900_E;
      END_IF

    // ANLEGEN ==================================================
    STEP_900_E:
      bpFehler := TRUE;

    // ANLEGEN ==================================================
    STEP_1000_E:
      bpDone := TRUE;

      IF ( starrStationBasisParameter[wStation].eStatusAuftrag = eAuftragErfolgreich ) THEN

        IF Auftragsdaten.bModell  OR NOT (starrStationBasisParameter[wStation].stMKs.stStationsOptionen.stGlastransport.bScheibenVermessen) THEN
          Auftragsdaten.wAuftrag := eStation_Warte_Auf_Austransport;
        ELSE
          Auftragsdaten.wAuftrag := eStation_Hoehenmessung;
        END_IF

      ELSIF ( starrStationBasisParameter[wStation].eStatusAuftrag = eAuftragWiederholen ) THEN
        steplSchritt := STEP_0_E;

      END_IF

  // ANLEGEN ==================================================
  END_CASE
END_IF

IF bpReset THEN
  blAktiv := FALSE;
  bpFehler := FALSE;
  bpReset := FALSE;
  bpDone := FALSE;
  steplSchritt := STEP_0_E;
  starrStationBasisParameter[wStation].bAnlegen := FALSE;
END_IF
END_FUNCTION_BLOCK
